(* IEC 61131-3 sources: daoli-st-library/DL_Algo (part 19) *)

(* ---- FB_DL_Q15BiquadFilter.st ---- *)
(*
  FB_DL_Q15BiquadFilter —— Q15 定点二阶 IIR 滤波：系数定点化、中间累加防溢出、移位饱和输出
  分类：DL_Algo | 复杂度：3 | 轮次：R86
  开源溯源：道莅原创（clean-room 自研，纯 IEC 61131-3 通用算法），无外部代码引用
  许可证：MIT

  职责：以直接 II 型转置（DF2T）结构实现二阶 IIR：y[n] = b0*x[n] + z1[n-1]；
        z1[n] = b1*x[n] - a1*y[n] + z2[n-1]；z2[n] = b2*x[n] - a2*y[n]。
        全部乘加在 DINT 内完成（Q15 × Q15 得 Q30），统一做「四舍五入右移 15 位 + Q15 饱和」，不调用任何外部库件。
  输入契约：arrCoef[0..4] = b0 / b1 / b2 / a1 / a2，均为 Q15 系数（±1.0 对应 ±32767）；
            iIn 为 Q15 输入；xReset 上升至真清历史；xEnable = FALSE 时清历史并输出 0。
  输出契约：iOut 为 Q15 输出；xOverflow 表示本拍发生了乘法累加或输出的饱和（信息级，可每拍重算）。
  边界：① 无除法、无开方，除零风险为零；② 所有移位用「乘 32768 / 除 32768」表达，避免方言 SHL/SHR 语义差异；
        ③ 定点饱和阈值 Q15_MAX / Q15_MIN 用 VAR CONSTANT 钉死；④ 零全局耦合、零物理地址、零库件依赖（R16）。
*)

FUNCTION_BLOCK FB_DL_Q15BiquadFilter
VAR_INPUT
    xEnable  : BOOL := TRUE;                              // 使能，FALSE 时清历史并输出零 [—] / Enable, false clears history
    xReset   : BOOL := FALSE;                             // 复位，真时清历史（单拍即可，无需沿） [—] / Reset, clears the history
    iIn      : INT  := 0;                                 // Q15 定点输入 [Q15] / The Q15 fixed point input
    arrCoef  : ARRAY[0..4] OF INT;                        // Q15 系数 b0/b1/b2/a1/a2 [Q15] / The Q15 coefficients
END_VAR
VAR_OUTPUT
    iOut      : INT;                                      // Q15 定点输出 [Q15] / The Q15 fixed point output
    xOverflow : BOOL;                                     // 本拍发生饱和（信息级） [—] / A saturation occurred this scan
END_VAR
VAR
    arrHist   : ARRAY[0..3] OF INT;                       // 历史：0=z1 1=z2 2=上拍输入 3=上拍输出 [Q15] / History slots
    diProd1   : DINT;                                     // 第一乘积项（Q30） [Q30] / The first product term
    diProd2   : DINT;                                     // 第二乘积项（Q30） [Q30] / The second product term
    diAcc     : DINT;                                     // 累加器（Q30） [Q30] / The Q30 accumulator
    diSh      : DINT;                                     // 四舍五入右移后的 Q15 暂存 [Q15] / The rounded Q15 stage
    diSum     : DINT;                                     // Q15 域饱和加法暂存 [Q15] / The Q15 domain saturating sum
    iNewZ1    : INT;                                      // 新的 z1 状态 [Q15] / The new z1 state
    iNewZ2    : INT;                                      // 新的 z2 状态 [Q15] / The new z2 state
    iSat      : INT;                                      // 饱和后的输出暂存 [Q15] / The saturated output stage
END_VAR
VAR CONSTANT
    Q15_MAX   : DINT := 32767;                            // Q15 上界 [-] / The Q15 upper bound
    Q15_MIN   : DINT := -32768;                           // Q15 下界 [-] / The Q15 lower bound
    DL_BQ_RND : DINT := 16384;                            // 右移 15 位的四舍五入偏置（2^14） [-] / The rounding bias
    DL_BQ_SC  : DINT := 32768;                            // Q15 定标因子（2^15） [-] / The Q15 scaling factor
    DL_BQ_Z   : DINT := 0;                                // 整型零常量 [Q15] / The integer zero constant
    DL_BQ_I0  : INT := 0;                                 // 整型零常量（INT 域） [Q15] / The integer zero constant in INT domain
    DL_BQ_I1  : INT := 1;                                 // 整型一常量（下标） [下标] / The integer one constant
    DL_BQ_I2  : INT := 2;                                 // 整型二常量（下标） [下标] / The integer two constant
    DL_BQ_I3  : INT := 3;                                 // 整型三常量（下标） [下标] / The integer three constant
    DL_BQ_I4  : INT := 4;                                 // 整型四常量（下标） [下标] / The integer four constant
END_VAR

// 段 1｜出口预置（本拍饱和标志每拍重算，属信息级）
xOverflow := FALSE;                                       // 饱和标志预置假 / preset the saturation flag false
iOut := DL_BQ_I0;                                         // 输出预置零 [Q15] / preset the output zero

// 段 2｜复位 / 失能闸：清全部历史并输出零（唯一复位路径）
IF xReset OR NOT xEnable THEN                             // 复位或失能 / reset asserted or disabled
    arrHist[DL_BQ_I0] := DL_BQ_I0;                        // z1 清零 [Q15] / clear z1
    arrHist[DL_BQ_I1] := DL_BQ_I0;                        // z2 清零 [Q15] / clear z2
    arrHist[DL_BQ_I2] := DL_BQ_I0;                        // 上拍输入清零 [Q15] / clear the previous input
    arrHist[DL_BQ_I3] := DL_BQ_I0;                        // 上拍输出清零 [Q15] / clear the previous output
    iOut := DL_BQ_I0;                                     // 输出零 [Q15] / output zero
    xOverflow := FALSE;                                   // 清饱和标志 [—] / clear the saturation flag
ELSE
    // 段 3｜y[n] = b0*x[n] + z1[n-1]（两项之和界内可证：|b0*x| <= 1.073e9，|z1*2^15| <= 1.073e9）
    diProd1 := INT_TO_DINT(arrCoef[DL_BQ_I0]) * INT_TO_DINT(iIn);          // b0*x [Q30] / b0 times x
    diProd2 := INT_TO_DINT(arrHist[DL_BQ_I0]) * DL_BQ_SC;                  // z1 左移 15 位 [Q30] / z1 scaled to Q30
    diAcc := diProd1 + diProd2;                                            // 两项求和 [Q30] / sum the two terms
    IF diAcc >= DL_BQ_Z THEN                                               // 非负做加偏置舍入 / non negative rounding
        diSh := (diAcc + DL_BQ_RND) / DL_BQ_SC;                            // 四舍五入右移 15 位 [Q15] / rounded shift right
    ELSE
        diSh := (diAcc - DL_BQ_RND) / DL_BQ_SC;                            // 负值做减偏置舍入 [Q15] / rounded shift right
    END_IF
    IF diSh > Q15_MAX THEN                                                 // 输出上越界 / the output exceeds the upper bound
        iSat := DINT_TO_INT(Q15_MAX);                                      // 饱和到 Q15_MAX [Q15] / saturate high
        xOverflow := TRUE;                                                 // 置饱和标志 [—] / raise the saturation flag
    ELSIF diSh < Q15_MIN THEN                                              // 输出下越界 / the output exceeds the lower bound
        iSat := DINT_TO_INT(Q15_MIN);                                      // 饱和到 Q15_MIN [Q15] / saturate low
        xOverflow := TRUE;                                                 // 置饱和标志 [—] / raise the saturation flag
    ELSE
        iSat := DINT_TO_INT(diSh);                                         // 界内直接转换 [Q15] / in range conversion
    END_IF
    iOut := iSat;                                                          // 本拍输出 [Q15] / the output of this scan

    // 段 4｜z1[n] = b1*x[n] - a1*y[n] + z2[n-1]（先算 Q30 两项差，再移位，再在 Q15 域饱和加 z2）
    diProd1 := INT_TO_DINT(arrCoef[DL_BQ_I1]) * INT_TO_DINT(iIn);          // b1*x [Q30] / b1 times x
    diProd2 := INT_TO_DINT(arrCoef[DL_BQ_I3]) * INT_TO_DINT(iSat);         // a1*y [Q30] / a1 times y
    diAcc := diProd1 - diProd2;                                            // 两项差（界内 |差| <= 2.147e9 可证） [Q30]
    IF diAcc >= DL_BQ_Z THEN                                               // 非负做加偏置舍入 / non negative rounding
        diSh := (diAcc + DL_BQ_RND) / DL_BQ_SC;                            // 四舍五入右移 15 位 [Q15] / rounded shift right
    ELSE
        diSh := (diAcc - DL_BQ_RND) / DL_BQ_SC;                            // 负值做减偏置舍入 [Q15] / rounded shift right
    END_IF
    diSum := diSh + INT_TO_DINT(arrHist[DL_BQ_I1]);                        // 加上 z2（|和| <= 98304 界内） [Q15] / add z2
    IF diSum > Q15_MAX THEN                                                // z1 上越界 / z1 exceeds the upper bound
        iNewZ1 := DINT_TO_INT(Q15_MAX);                                    // 饱和到 Q15_MAX [Q15] / saturate high
        xOverflow := TRUE;                                                 // 置饱和标志 [—] / raise the saturation flag
    ELSIF diSum < Q15_MIN THEN                                             // z1 下越界 / z1 exceeds the lower bound
        iNewZ1 := DINT_TO_INT(Q15_MIN);                                    // 饱和到 Q15_MIN [Q15] / saturate low
        xOverflow := TRUE;                                                 // 置饱和标志 [—] / raise the saturation flag
    ELSE
        iNewZ1 := DINT_TO_INT(diSum);                                      // 界内直接转换 [Q15] / in range conversion
    END_IF

    // 段 5｜z2[n] = b2*x[n] - a2*y[n]（同段 4 的判溢出 + 舍入 + 饱和口径）
    diProd1 := INT_TO_DINT(arrCoef[DL_BQ_I2]) * INT_TO_DINT(iIn);          // b2*x [Q30] / b2 times x
    diProd2 := INT_TO_DINT(arrCoef[DL_BQ_I4]) * INT_TO_DINT(iSat);         // a2*y [Q30] / a2 times y
    diAcc := diProd1 - diProd2;                                            // 两项差 [Q30] / the difference of the two terms
    IF diAcc >= DL_BQ_Z THEN                                               // 非负做加偏置舍入 / non negative rounding
        diSh := (diAcc + DL_BQ_RND) / DL_BQ_SC;                            // 四舍五入右移 15 位 [Q15] / rounded shift right
    ELSE
        diSh := (diAcc - DL_BQ_RND) / DL_BQ_SC;                            // 负值做减偏置舍入 [Q15] / rounded shift right
    END_IF
    IF diSh > Q15_MAX THEN                                                 // z2 上越界 / z2 exceeds the upper bound
        iNewZ2 := DINT_TO_INT(Q15_MAX);                                    // 饱和到 Q15_MAX [Q15] / saturate high
        xOverflow := TRUE;                                                 // 置饱和标志 [—] / raise the saturation flag
    ELSIF diSh < Q15_MIN THEN                                              // z2 下越界 / z2 exceeds the lower bound
        iNewZ2 := DINT_TO_INT(Q15_MIN);                                    // 饱和到 Q15_MIN [Q15] / saturate low
        xOverflow := TRUE;                                                 // 置饱和标志 [—] / raise the saturation flag
    ELSE
        iNewZ2 := DINT_TO_INT(diSh);                                       // 界内直接转换 [Q15] / in range conversion
    END_IF

    // 段 6｜状态统一提交（两段式：先算新值后写回，避免同拍读写串扰）
    arrHist[DL_BQ_I2] := iIn;                                             // 记录上拍输入 [Q15] / record the previous input
    arrHist[DL_BQ_I3] := iSat;                                            // 记录上拍输出 [Q15] / record the previous output
    arrHist[DL_BQ_I0] := iNewZ1;                                          // 提交新的 z1 [Q15] / commit z1
    arrHist[DL_BQ_I1] := iNewZ2;                                          // 提交新的 z2 [Q15] / commit z2
END_IF
END_FUNCTION_BLOCK

(* ---- FB_DL_QuantizeFilter.st ---- *)
(*==============================================================================
 * 组件名称 (Component)  : FB_DL_QuantizeFilter
 * 所属子库 (Sublibrary) : DL_Algo
 * 当前版本 (Version)    : 1.0.0
 * 兼容性   (Platform)   : CODESYS 3.5+ / TwinCAT 3 / 汇川 InoProShop / 施耐德 Machine Expert
 *                         仅依赖 Standard.library（ROUND / ABS），零厂商私有库
 * 功能描述 (Function)   : **量化取整 + 回差防抖**（有状态件）。
 *                         第一步量化：fQ := ROUND(fIn / fStep) × fStep（就近取整到步距倍数）；
 *                         第二步回差：仅当 |fQ - fOut| > fHyst 时才把 fOut 更新为 fQ，
 *                         否则保持。两步合起来解决「量化值在相邻两档之间反复跳」的现场顽症
 *                         （典型：0.5 单位步距的设定值显示与控制字抖动）。
 *                         与无状态取整 FC（FC_DL_QuantizeStep）的差别：那件每拍直接输出
 *                         量化值、无记忆；本件带上一档记忆与回差，切换次数显著下降。
 * 接口     (Interface)  : 输入 bEnable 使能、bReset 复位到当前量化值、fIn 采样输入 [EU]、
 *                         fStep 量化步距（必须 > 0） [EU]、fHyst 切换回差（>= 0） [EU]；
 *                         输出 fOut 量化并防抖后的输出 [EU]、fQuantized 原始量化值（诊断） [EU]、
 *                         bUpdated 本拍是否切换档位、bValid 输出有效、bError、uErrorId。
 * 边界     (Boundary)   : ① 属主边界：只做步距量化与回差防抖，不做死区保持（另件）、不做限速（另件）。
 *                         ② **除零防护（R4 硬要求）**：fStep 参与除法 fIn / fStep，
 *                         必须先判 fStep > 0，否则故障级 16#0009_0003，输出冻结。
 *                         fStep = 0 不允许「静默当直通」，否则调用方看不出配置错误。
 *                         ③ fHyst < 0 → 故障级 16#0009_0003（负回差等于放大抖动）。
 *                         ④ 非有限防御：fIn / fStep / fHyst 三个浮点入参逐一枚举。
 *                         ⑤ 取整一律用 ROUND（禁止 TRUNC(x)+1 这类手工进位）。
 *                         ⑥ 恢复路径：bEnable=FALSE 或 bReset=TRUE 解除故障态。
 *                         ⑦ 零全局耦合（无 GVL / VAR_EXTERNAL / 物理地址）。
 * 分工声明 (Scope)      : 与无状态 `FC_DL_QuantizeStep` 分工：单拍取整归那件、
 *                         带记忆的回差防抖归本件；与 `FB_DL_DeadbandFilter` 分工：
 *                         连续量死区归那件、离散档位回差归本件。
 * 来源标签 (Source Tag) : 原创实现（无外部代码引入）
 * 码表     (Codes)      : 16#0009_0000 无故障 / 16#0009_0002 入参非有限（故障级）/
 *                         16#0009_0003 步距或回差非法（故障级）/ 16#0009_0005 非法状态（故障级）。
 * 红线自检 (Redline)    : R1 ✓ 零 GVL/VAR_EXTERNAL ｜ R2 ✓ 零 %I/%Q/%M ｜ R3 ✓ 纯 IEC 61131-3
 *                         R4 ✓ 步距前置判零（除零防护）+ 三浮点入参非有限判 + ROUND 取整 ｜ R5 ✓ 声明逐行同行双语注释
 *                         R6 ✓ 四态 ENUM + CASE + ELSE 兜底 ｜ R7 N/A（无 TON / 边沿实例）
 * 修订历史 (Revision)   : 2026-11-23  v1.0.0  R77 首版（批次 B3 · 序号 15）
 * 验收向量 (Acceptance) : ① fStep=0.5, fHyst=0.2, fIn=1.24 → fQ=ROUND(2.48)×0.5=2×0.5=1.0，
 *                         |1.0 - fOut(初 0)|=1.0 > 0.2 → fOut=1.0, bUpdated=TRUE；
 *                         ② 随后 fIn=1.26 → fQ=ROUND(2.52)×0.5=3×0.5=1.5，|1.5-1.0|=0.5 > 0.2 → fOut=1.5；
 *                         ③ 随后 fIn=1.30 → fQ=1.5，|1.5-1.5|=0 <= 0.2 → fOut 保持 1.5, bUpdated=FALSE；
 *                         ④ fStep=0.0 → uErrorId=16#0009_0003，bError=TRUE（不静默直通）；
 *                         ⑤ fHyst=-0.1 → uErrorId=16#0009_0003，bError=TRUE。
 *==============================================================================*)

(*-----------------------------------------------------------------------------
 * 枚举: E_DL_QuantState（量化防抖状态机，归属 DL_Algo，与本件同文件，全库唯一属主）
 *----------------------------------------------------------------------------*)
TYPE E_DL_QuantState :
(
    eInit  := 0,    // 首扫 / 复位后：输出直取当前量化值 / First scan or after reset: output equals quantized value
    eRun   := 10,   // 运行态：量化 + 回差判定 / Running: quantize plus hysteresis decision
    eHold  := 20,   // 保持态：未使能，输出冻结 / Hold: disabled, output frozen
    eFault := 99    // 故障态：输出冻结，等待 bEnable 跌落或 bReset / Fault: frozen until cleared
);
END_TYPE

FUNCTION_BLOCK FB_DL_QuantizeFilter
VAR_INPUT
    bEnable : BOOL := FALSE;   // 使能，FALSE 冻结输出 / Enable, FALSE freezes output
    bReset  : BOOL := FALSE;   // 复位到当前量化值（单拍有效） / Reset to current quantized value, single scan
    fIn     : LREAL := 0.0;    // 采样输入 [EU] / Sampling input [EU]
    fStep   : LREAL := 1.0;    // 量化步距，必须 > 0 [EU] / Quantisation step, must be positive [EU]
    fHyst   : LREAL := 0.0;    // 切换回差，必须 >= 0 [EU] / Switching hysteresis, must be non-negative [EU]
END_VAR
VAR_OUTPUT
    fOut       : LREAL;   // 量化并防抖后的输出 [EU] / Quantised and debounced output [EU]
    fQuantized : LREAL;   // 原始量化值（诊断用） [EU] / Raw quantised value for diagnostics [EU]
    bUpdated   : BOOL;    // 本拍是否切换档位 [-] / Whether the output switched this scan
    bValid     : BOOL;    // 输出有效标志 [-] / Output valid flag
    bError     : BOOL;    // 故障标志，与 uErrorId 联动 [-] / Fault flag coupled with uErrorId
    uErrorId   : UDINT;   // 故障码，0 = 无故障 [-] / Error code, zero means healthy
END_VAR
VAR
    _bNonFin : BOOL;              // 入参非有限标志 [-] / Non-finite input flag
    _fRatio  : LREAL;             // 步距倍数（取整前） [-] / Step multiple before rounding
    eState   : E_DL_QuantState;   // 状态机当前状态 [-] / Current state
END_VAR
VAR CONSTANT
    DL_QTF_ZERO : LREAL := 0.0;   // 零基准（含非有限判零） [-] / Zero base including non-finite probe
END_VAR

(* —— 段 1：非有限防御（fIn / fStep / fHyst 三入参逐一枚举） —— *)
uErrorId := 16#0009_0000;                          // 预置无故障 / Preset healthy
_bNonFin := (fIn <> fIn) OR ((fIn - fIn) <> DL_QTF_ZERO);            // 输入非有限 / Input non-finite
_bNonFin := _bNonFin OR (fStep <> fStep) OR ((fStep - fStep) <> DL_QTF_ZERO);   // 步距非有限
_bNonFin := _bNonFin OR (fHyst <> fHyst) OR ((fHyst - fHyst) <> DL_QTF_ZERO);   // 回差非有限
IF _bNonFin THEN
    eState   := eFault;                            // 强制故障态 / Force fault state
    uErrorId := 16#0009_0002;                      // 故障级：入参非有限 / Fault: non-finite input
END_IF

(* —— 段 2：步距与回差域闸（步距必须严格正：它是除数；回差必须非负） —— *)
IF (fStep <= DL_QTF_ZERO) OR (fHyst < DL_QTF_ZERO) THEN
    eState   := eFault;                            // 参数非法进故障态 / Illegal parameter goes to fault
    uErrorId := 16#0009_0003;                      // 故障级：步距或回差非法 / Fault: illegal step or hysteresis
    fQuantized := DL_QTF_ZERO;                     // 诊断量回 0 / Diagnostic value zeroed
END_IF

(* —— 段 3：复位请求 → 回首扫 —— *)
IF bReset THEN
    eState := eInit;
END_IF

(* —— 段 4：状态派生 —— *)
IF NOT bEnable THEN
    eState := eHold;                               // 未使能：冻结 / Disabled: freeze
ELSIF eState = eFault THEN
    eState := eFault;                              // 故障态保持 / Fault holds
ELSIF eState = eInit THEN
    eState := eInit;                               // 首扫保持一拍 / Init holds one scan
ELSE
    eState := eRun;
END_IF

(* —— 段 5：主状态机（CASE 覆盖 + ELSE 兜底） —— *)
CASE eState OF

    eInit:
        _fRatio     := fIn / fStep;                // 步距倍数（fStep 已在段 2 判正） / Step multiple, step proven positive
        fQuantized  := ROUND(_fRatio) * fStep;     // 就近量化（禁止 TRUNC+1 手工进位） / Nearest quantisation
        fOut        := fQuantized;                 // 首拍直取量化值 / First scan adopts quantised value
        bUpdated    := TRUE;
        bValid      := TRUE;
        eState      := eRun;

    eRun:
        _fRatio    := fIn / fStep;                 // 步距倍数 / Step multiple
        fQuantized := ROUND(_fRatio) * fStep;      // 就近量化 / Nearest quantisation
        IF ABS(fQuantized - fOut) > fHyst THEN
            fOut     := fQuantized;                // 超出回差：切换档位 / Beyond hysteresis: switch
            bUpdated := TRUE;
        ELSE
            (* 回差内：保持原档位，避免相邻档反复跳变 / Inside hysteresis: hold current step *)
            bUpdated := FALSE;
        END_IF
        bValid := TRUE;

    eHold:
        (* 未使能：输出、量化诊断值、切换标志全部冻结 / Disabled: output, diagnostic and flag frozen *)
        bUpdated := FALSE;
        bValid   := FALSE;

    eFault:
        (* 故障态：输出冻结保持上拍值（不推 0，避免下游误判） / Fault: output frozen *)
        bUpdated := FALSE;
        bValid   := FALSE;

    ELSE
        eState     := eFault;
        bUpdated   := FALSE;
        bValid     := FALSE;
        fQuantized := DL_QTF_ZERO;
        uErrorId   := 16#0009_0005;                // 故障级：非法状态 / Fault: illegal state

END_CASE;

(* —— 段 6：出口映射（bError 与 uErrorId 同源；本件无信息级码） —— *)
bError := (uErrorId <> 16#0009_0000);

END_FUNCTION_BLOCK

(* ---- FB_DL_RampGenerator.st ---- *)
(*==============================================================================
 * 组件名称 (Component)  : FB_DL_RampGenerator
 * 所属子库 (Sublibrary) : DL_Algo
 * 当前版本 (Version)    : 1.0.1
 * 兼容性   (Platform)   : CODESYS 3.5 / TwinCAT 3 / 汇川 InoProShop / Machine Expert
 *                         仅依赖 Standard.library（LIMIT / MIN / ABS / SIGN），零厂商方言
 * 功能描述 (Function)   : 线性设定值斜坡发生器。把阶跃目标值变为按独立上升/下降
 *                         速率（EU/s）平滑逼近的斜坡输出，防止操作员大阶跃直接
 *                         冲击执行器。支持暂停保持（bHold 冻结当前值）与跟踪回投
 *                         （bTrack + fTrackValue 投切无扰动）。
 *                         斜率为 0 表示该方向冻结（保持输出，绝不直通，防误操作）。
 *                         到达判定以限幅后的实际输出为准，防止目标超量程时死等。
 * 开源溯源 (Origin)     : 原创实现。算法思想源自 IEC 61131-3 标准函数语义与
 *                         PLCopen Coding Guidelines 的周期安全约定，
 *                         未复制任何厂商私有库源码。
 * 本文件内含       : TYPE  E_DL_RampState（配套枚举，归属 DL_Algo）
 *                    FB    FB_DL_RampGenerator
 * 依赖     (Depends)    : 无 DL_ 内部依赖；Standard.library: LIMIT / MIN / ABS / SIGN
 * 红线自检 (Redline)    : R1 ✓ 零全局变量表与外部变量引用 ｜ R2 ✓ 零物理 IO 地址直写
 *                         R3 ✓ 纯 IEC 61131-3 ｜ R4 ✓ 速率/量程钳位+非有限值拒绝
 *                         R5 ✓ 全变量中英双语同行注释 ｜ R6 ✓ 六态 ENUM+CASE+ELSE
 *                         R7 N/A（无定时器/边沿实例）
 * 【边界披露 / Boundary disclosure】
 *   B1 速率 <= 0 视为非法：置 16#0002_0601 且该方向步长为 0（冻结），绝不直通。
 *   B2 目标非有限值（NaN 或幅值超 1.0E30）：本拍拒绝更新，保持上一拍输出。
 *   B3 rOutMin > rOutMax：自动对调并置 16#0002_0001，不中断扫描。
 *   B4 目标超量程不截断目标，仅限幅输出；到达判定用限幅后实际值，防死等。
 * 【验收向量 / Acceptance vectors】
 *   V1  fTarget 0→100，fRateUp=10 EU/s，tSampleTime=T#100MS → 每拍 +1.0 EU，
 *       10 s 后 fOut≈100、bDone=TRUE
 *   V2  fTarget 100→30，fRateDown=10 EU/s → 每拍 -1.0 EU、bMoving=TRUE
 *   V3  bHold=TRUE → fOut 冻结、状态 eHold；释放后继续逼近目标
 *   V4  fRateUp=0 → 16#0002_0601，向上移动冻结、fOut 保持
 *   V5  bTrack 一拍（fTrackValue=50）→ fOut=50，下一拍从 50 继续斜坡（无扰动）
 *   V6  rOutMin=100 > rOutMax=0 → 自动对调、16#0002_0001
 *   V7  fTarget=NaN → 16#0002_0004，fOut 保持上一拍值
 * 修订历史 (Revision)   :
 *   2026-11-15  v1.0.0  首版入库（Round 04 · Phase 3 · DL_Algo 批次）
 *   2026-11-15  v1.0.1  阶段五终审精修：首扫自动跟踪判据修复（bInit 判据
 *                       反向导致首扫不跟踪），对齐通用约定 0-6
 *============================================================================*)

(*-----------------------------------------------------------------------------
 * 枚举: E_DL_RampState（归属 DL_Algo，与 FB_DL_RampGenerator 同文件）
 * 含义: 斜坡状态机离散状态。数值步长留空位便于后续插态而不破坏已有工程。
 *----------------------------------------------------------------------------*)
TYPE E_DL_RampState :
(
    eIdle    := 0,    // 空闲态：未使能或等待评估，输出保持 / Idle state, output frozen
    eHold    := 10,   // 暂停保持态：操作员请求冻结当前输出 / Hold state, output frozen on operator request
    eRampUp  := 20,   // 上升斜坡态：按 fRateUpEff 步进逼近目标 / Ramping up with effective up rate
    eRampDown:= 30,   // 下降斜坡态：按 fRateDownEff 步进逼近目标 / Ramping down with effective down rate
    eDone    := 40,   // 到达态：输出与目标偏差在容差内 / Done state, deviation within tolerance
    eFault   := 99    // 故障兜底态：非法状态拦截，自动回空闲 / Fault fallback, auto recover to idle
);
END_TYPE

(*==============================================================================
 * 功能块: FB_DL_RampGenerator
 * 调用约定: 每个扫描周期无条件调用一次；bTrack 使能时输出立即跟随 fTrackValue。
 * 无状态泄漏: 全部状态驻留于实例私有 VAR，可多实例并行互不影响。
 * 速率披露: 输出相对目标的延迟 = 偏差量 / 对应方向速率（线性，非固定时间）。
 *============================================================================*)
FUNCTION_BLOCK FB_DL_RampGenerator
VAR_INPUT
    bEnable     : BOOL := FALSE;        // 使能标志，FALSE 时斜坡停止并保持输出 / Enable flag, FALSE stops ramp and holds output
    fTarget     : REAL := 0.0;          // 目标值 [EU]，可为任意有限值 / Target value [EU], any finite value
    fRateUp     : REAL := 10.0;         // 上升速率 [EU/s]，<=0 视为非法冻结 / Up rate [EU/s], <=0 illegal and frozen
    fRateDown   : REAL := 10.0;         // 下降速率 [EU/s]，<=0 视为非法冻结 / Down rate [EU/s], <=0 illegal and frozen
    bHold       : BOOL := FALSE;        // 暂停保持请求，TRUE 冻结在当前值 / Hold request, TRUE freezes at current value
    bTrack      : BOOL := FALSE;        // 跟踪使能，TRUE 时输出立即跟随 fTrackValue / Track enable, output follows fTrackValue instantly
    fTrackValue : REAL := 0.0;          // 跟踪值 [EU]，投切无扰动基准 / Track value [EU], bumpless transfer reference
    rOutMin     : REAL := -1.0E10;      // 输出下限 [EU]，大于上限时自动对调 / Output lower limit [EU], swapped if greater
    rOutMax     : REAL := 1.0E10;       // 输出上限 [EU]，小于下限时自动对调 / Output upper limit [EU], swapped if smaller
    tSampleTime : TIME := T#100MS;      // 采样周期 [s]，小于 10ms 钳位为 10ms / Sample time [s], clamped to 10ms minimum
END_VAR
VAR_OUTPUT
    fOut        : REAL;                 // 斜坡输出 [EU] / Ramp output [EU]
    bDone       : BOOL;                 // 到达目标标志：偏差在容差内 / Done flag, deviation within tolerance
    bMoving     : BOOL;                 // 斜坡进行中标志 / Ramp in progress flag
    fRemain     : REAL;                 // 距目标剩余量 [EU] = fTarget - fOut / Remaining amount to target [EU]
    bError      : BOOL;                 // 故障标志（瞬时，逐拍重算） / Fault flag, transient, recomputed every scan
    uErrorId    : UDINT;                // 故障码，0 = 无故障 / Error code, 0 = no error
END_VAR
VAR
    fRateUpEff  : REAL;                 // 钳位后的有效上升速率 [EU/s] / Effective clamped up rate [EU/s]
    fRateDownEff: REAL;                 // 钳位后的有效下降速率 [EU/s] / Effective clamped down rate [EU/s]
    fDt         : REAL;                 // 折算后的采样周期 [s] / Converted sample period [s]
    fDelta      : REAL;                 // 本拍目标与输出的偏差 [EU] / Deviation between target and output [EU]
    fStep       : REAL;                 // 本拍允许的最大步长 [EU] / Max step allowed this scan [EU]
    bTgtValid   : BOOL;                 // 目标为有限值的合法性标志 / Target finite validity flag
    bInit       : BOOL;                 // 首扫标志：首扫自动跟踪 fTrackValue / First scan flag, auto track on first scan
    eState      : E_DL_RampState;       // 主状态机当前状态 / Current state of the main state machine
END_VAR
VAR CONSTANT
    DL_RAMP_EPS     : REAL := 1.0E-6;   // 到达判定容差 [EU]，浮点差值比较 / Arrival tolerance [EU], float diff compare
    DL_RAMP_RATE_MAX: REAL := 1.0E10;   // 速率上限钳位 [EU/s]，防溢出 / Rate upper clamp [EU/s], overflow guard
END_VAR

(*------------------------------------------------------------------------------
 * 段 1｜公共参数处理（通用约定 0-1/0-2/0-3）：周期钳位、量程对调、故障码瞬时清零
 *      Common parameter handling: sample time clamp, limit swap, transient code reset
 *-----------------------------------------------------------------------------*)
uErrorId := 16#0000_0000;               // 故障码逐拍重算（瞬时语义） / Error code recomputed every scan
bError   := FALSE;                      // 故障标志逐拍重算 / Fault flag recomputed every scan

IF tSampleTime < T#10MS THEN
    fDt      := TIME_TO_REAL(T#10MS) / 1000.0; // 非法周期钳位为 10ms / Illegal period clamped to 10ms
    uErrorId := 16#0002_0002;           // 采样周期非法已钳位 / Sample time illegal, clamped
ELSE
    fDt      := TIME_TO_REAL(tSampleTime) / 1000.0; // 周期换算为秒 [s] / Period converted to seconds [s]
END_IF

IF rOutMin > rOutMax THEN
    fOut := LIMIT(rOutMax, fOut, rOutMin); // 对调后按新序限幅输出 / Clamp output with swapped limits
    uErrorId := 16#0002_0001;           // 参数越界已对调 / Limits out of order, swapped
ELSE
    fOut := LIMIT(rOutMin, fOut, rOutMax); // 正常序限幅输出 / Clamp output with normal limits
END_IF

(*------------------------------------------------------------------------------
 * 段 2｜速率钳位：<=0 非法（冻结方向），超上限钳位（边界 B1）
 *      Rate clamping: <=0 illegal (freeze direction), over-limit clamped
 *-----------------------------------------------------------------------------*)
IF fRateUp <= 0.0 THEN
    fRateUpEff := 0.0;                  // 非法速率冻结为 0，步长为 0 / Illegal rate frozen to zero step
    uErrorId   := 16#0002_0601;         // 速率非法已钳位 / Rate illegal, clamped
ELSIF fRateUp > DL_RAMP_RATE_MAX THEN
    fRateUpEff := DL_RAMP_RATE_MAX;     // 超上限钳位防溢出 / Over-limit clamped for overflow guard
    uErrorId   := 16#0002_0601;         // 速率非法已钳位 / Rate illegal, clamped
ELSE
    fRateUpEff := fRateUp;              // 合法速率直通 / Valid rate passed through
END_IF

IF fRateDown <= 0.0 THEN
    fRateDownEff := 0.0;                // 非法速率冻结为 0，步长为 0 / Illegal rate frozen to zero step
    uErrorId     := 16#0002_0601;       // 速率非法已钳位 / Rate illegal, clamped
ELSIF fRateDown > DL_RAMP_RATE_MAX THEN
    fRateDownEff := DL_RAMP_RATE_MAX;   // 超上限钳位防溢出 / Over-limit clamped for overflow guard
    uErrorId     := 16#0002_0601;       // 速率非法已钳位 / Rate illegal, clamped
ELSE
    fRateDownEff := fRateDown;          // 合法速率直通 / Valid rate passed through
END_IF

(*------------------------------------------------------------------------------
 * 段 3｜目标合法性判定（边界 B2）：非有限值本拍拒绝，保持上一拍目标行为
 *      Target validity: non-finite value rejected this scan, previous behavior kept
 *-----------------------------------------------------------------------------*)
bTgtValid := NOT (fTarget <> fTarget) AND (ABS(fTarget) <= 1.0E30); // NaN 判别 + 幅值防御 / NaN check plus magnitude guard
IF NOT bTgtValid THEN
    uErrorId := 16#0002_0004;           // 输入非有限值已拒绝 / Non-finite input rejected
END_IF

(*------------------------------------------------------------------------------
 * 段 4｜跟踪与首扫（通用约定 0-6）：投切无扰动，首扫自动跟踪 fTrackValue
 *      Tracking and first scan: bumpless transfer, first scan auto track
 *-----------------------------------------------------------------------------*)
IF bTrack OR (NOT bInit) THEN
    fOut   := LIMIT(rOutMin, fTrackValue, rOutMax); // 输出立即跟随跟踪值 / Output follows track value instantly
    eState := eIdle;                    // 回空闲重新评估方向 / Back to idle for direction re-evaluation
    bInit  := TRUE;                     // 首扫标志置位 / First scan flag set
END_IF

(*------------------------------------------------------------------------------
 * 段 5｜主状态机（红线 R6）：ENUM + CASE + ELSE 兜底
 *      Main state machine: ENUM + CASE with mandatory ELSE fallback
 *-----------------------------------------------------------------------------*)
fDelta := fTarget - fOut;               // 本拍偏差 [EU] / Deviation this scan [EU]

IF NOT bEnable THEN
    eState := eIdle;                    // 未使能：强制空闲、输出保持 / Disabled: force idle, output held
ELSE
    CASE eState OF

        eIdle:  // 空闲态：使能后按偏差方向选择迁移 / Idle: pick transition by deviation direction
            IF bTgtValid AND ABS(fDelta) > DL_RAMP_EPS THEN
                IF bHold THEN
                    eState := eHold;    // 保持请求优先 / Hold request has priority
                ELSIF fDelta > 0.0 THEN
                    eState := eRampUp;  // 目标在上方，进入上升 / Target above, ramp up
                ELSE
                    eState := eRampDown; // 目标在下方，进入下降 / Target below, ramp down
                END_IF
            ELSIF bTgtValid THEN
                eState := eDone;        // 已在容差内，直接到达 / Already within tolerance, done
            END_IF

        eHold:  // 暂停保持态：冻结输出直到释放 / Hold: freeze output until released
            IF NOT bHold THEN
                IF ABS(fDelta) <= DL_RAMP_EPS THEN
                    eState := eDone;    // 保持期间目标已到达 / Target reached during hold
                ELSIF fDelta > 0.0 THEN
                    eState := eRampUp;  // 释放后继续上升 / Resume ramp up after release
                ELSE
                    eState := eRampDown; // 释放后继续下降 / Resume ramp down after release
                END_IF
            END_IF

        eRampUp:  // 上升斜坡态：步长 = MIN(偏差, 速率*周期) / Ramp up: step = MIN(deviation, rate*period)
            IF ABS(fDelta) <= DL_RAMP_EPS THEN
                eState := eDone;        // 到达目标 / Target reached
            ELSIF fDelta < 0.0 THEN
                eState := eRampDown;    // 目标反转为下方 / Target switched below
            ELSIF bHold THEN
                eState := eHold;        // 保持请求 / Hold request
            ELSE
                fStep := MIN(fDelta, fRateUpEff * fDt); // 本拍步长 [EU] / Step this scan [EU]
                fOut  := fOut + fStep;  // 逐步逼近目标 / Step toward target
            END_IF

        eRampDown:  // 下降斜坡态：对称逻辑 / Ramp down: symmetric logic
            IF ABS(fDelta) <= DL_RAMP_EPS THEN
                eState := eDone;        // 到达目标 / Target reached
            ELSIF fDelta > 0.0 THEN
                eState := eRampUp;      // 目标反转为上方 / Target switched above
            ELSIF bHold THEN
                eState := eHold;        // 保持请求 / Hold request
            ELSE
                fStep := MIN(-fDelta, fRateDownEff * fDt); // 本拍步长 [EU] / Step this scan [EU]
                fOut  := fOut - fStep;  // 逐步逼近目标 / Step toward target
            END_IF

        eDone:  // 到达态：监视新目标 / Done: watch for new target
            IF bTgtValid AND ABS(fDelta) > DL_RAMP_EPS THEN
                IF bHold THEN
                    eState := eHold;    // 保持请求 / Hold request
                ELSIF fDelta > 0.0 THEN
                    eState := eRampUp;  // 新目标在上方 / New target above
                ELSE
                    eState := eRampDown; // 新目标在下方 / New target below
                END_IF
            END_IF

        eFault:  // 故障兜底态：无复位引脚，当拍回空闲重评，避免永久锁死 / Fault fallback: no reset pin, recover to idle
            eState := eIdle;            // 自动恢复空闲 / Auto recover to idle

        ELSE  // 非法状态拦截：任何未定义状态一律进故障态并置码 / Illegal state interception
            eState   := eFault;         // 强制故障态 / Force fault state
            uErrorId := 16#0002_0005;   // 非法状态兜底 / Illegal state fallback
            bError   := TRUE;           // 故障标志置位 / Fault flag set

    END_CASE;
END_IF

(*------------------------------------------------------------------------------
 * 段 6｜输出整形与状态引脚：限幅后实际值判定到达（边界 B4 防死等）
 *      Output shaping and status pins: arrival judged on clamped actual output
 *-----------------------------------------------------------------------------*)
IF rOutMin > rOutMax THEN
    fOut := LIMIT(rOutMax, fOut, rOutMin); // 对调序限幅（与段 1 一致） / Clamp with swapped order
ELSE
    fOut := LIMIT(rOutMin, fOut, rOutMax); // 正常序限幅 / Clamp with normal order
END_IF

fDelta  := fTarget - fOut;              // 限幅后重算偏差 [EU] / Deviation recomputed after clamping
fRemain := fDelta;                      // 距目标余量 [EU] / Remaining to target [EU]

bDone   := bEnable AND bTgtValid AND (ABS(fDelta) <= DL_RAMP_EPS); // 到达标志 / Done flag
bMoving := bEnable AND bTgtValid AND (NOT bHold)
           AND (ABS(fDelta) > DL_RAMP_EPS)
           AND ((eState = eRampUp) OR (eState = eRampDown));        // 斜坡进行中 / Ramp in progress
END_FUNCTION_BLOCK

(* ---- FB_DL_RateLimiter.st ---- *)
(*==============================================================================
 * 组件名称 (Component)  : FB_DL_RateLimiter
 * 所属子库 (Sublibrary) : DL_Algo
 * 当前版本 (Version)    : 1.0.0
 * 兼容性   (Platform)   : CODESYS 3.5 / TwinCAT 3 / 汇川 InoProShop / Machine Expert
 *                         仅依赖纯 IEC 61131-3 数学运算，零库依赖，零厂商方言
 * 功能描述 (Function)   : 变化率限制器（对应变化率限制语义）。输入阶跃时输出
 *                         以最大速率跟随，保护加热元件 / 执行器免受给定值阶跃
 *                         冲击；上升与下降速率独立可调，速率为 0 表示该方向不
 *                         限速直通（沿测量库惯例），负值非法按 0 处理并置码；
 *                         支持跟踪回投与限速进行中标志。
 * 开源溯源 (Origin)     : 原创实现。功能分类与参数域参考测量函数库中变化率
 *                         限制单元的公开语义描述，未复制任何厂商源码，
 *                         clean-room 重写。
 * 本文件内含       : TYPE  E_DL_RateState（配套枚举，归属 DL_Algo）
 *                    FB    FB_DL_RateLimiter
 * 依赖     (Depends)    : 无 DL_ 内部依赖；Standard.library 无实例依赖
 * 红线自检 (Redline)    : R1 ✓ 零全局变量表与外部变量引用 ｜ R2 ✓ 零物理 IO 地址直写
 *                         R3 ✓ 纯 IEC 61131-3 ｜ R4 ✓ 防除零+钳位+非有限值防御
 *                         R5 ✓ 全变量中英双语同行注释 ｜ R6 ✓ 五态 ENUM+CASE+ELSE
 *                         R7 ✓ 本块无定时器 / 边沿实例（无可刷新项，天然合规）
 * 修订历史 (Revision)   :
 *   2026-11-15  v1.0.0  首版入库 · Round 04 · Level 1 DL_Algo
 * 验收向量 (Acceptance) :
 *   V1 上升限速：fRateUp=10 EU/s, 输入阶跃 +100 → 输出每拍 +1 EU（100 ms 周期）
 *   V2 下降限速：fRateDown=5 EU/s, 输入阶跃 -100 → 输出每拍 -0.5 EU
 *   V3 零速率直通：fRateUp=0 → 上升方向立即跟随输入
 *   V4 到达直通：输出追上输入后 bLimiting=FALSE 且输出等于输入
 *   V5 跟踪：bTrack 置位 → 输出立即等于 fTrackValue
 *   V6 非有限值：输入写非法浮点 → 输出保持上一拍且码 0002_0004
 *============================================================================*)

(*-----------------------------------------------------------------------------
 * 枚举: E_DL_RateState（归属 DL_Algo，与 FB_DL_RateLimiter 同文件）
 * 含义: 变化率限制离散状态。数值步长留空位便于后续插态而不破坏已有工程。
 *----------------------------------------------------------------------------*)
TYPE E_DL_RateState :
(
    eIdle      := 0,   // 使能关：输出直通输入 / Idle: enable off, output follows input
    eFollow    := 10,  // 不限速直通：两方向均无需限速 / Follow: no rate limit needed in either direction
    eLimitUp   := 20,  // 上升限速：输出按最大上升速率逼近 / Limit up: output approaches at max rise rate
    eLimitDown := 30,  // 下降限速：输出按最大下降速率逼近 / Limit down: output approaches at max fall rate
    eFault     := 99   // 故障兜底态：非法状态进入，输出保持 / Fault fallback: illegal state, output held
);
END_TYPE

(*==============================================================================
 * 功能块: FB_DL_RateLimiter
 * 调用约定: 每个扫描周期无条件调用一次；采样周期引脚按子库通用约定配置。
 * 无状态泄漏: 全部状态驻留于实例私有 VAR，零全局引用，可多实例并行。
 * 工程披露: 输出变量自身即斜坡历史状态，不另设历史缓冲；实际变化率按本拍
 *           输出增量除以采样周期计算，供 HMI 趋势与诊断。
 *============================================================================*)
FUNCTION_BLOCK FB_DL_RateLimiter
VAR_INPUT
    bEnable     : BOOL := FALSE;      // 总使能，FALSE 时输出直通输入 / Master enable, FALSE passes input through
    fIn         : REAL := 0.0;        // 输入信号 [EU] / Input signal in engineering units
    fRateUp     : REAL := 0.0;        // 最大上升速率 [EU/s]，0 = 不限 / Max rising rate, 0 = unlimited
    fRateDown   : REAL := 0.0;        // 最大下降速率 [EU/s]，0 = 不限 / Max falling rate, 0 = unlimited
    bTrack      : BOOL := FALSE;      // 跟踪使能，TRUE 时输出立即跟随跟踪值 / Track enable, output follows track value
    fTrackValue : REAL := 0.0;        // 跟踪值 [EU]，用于无扰投切 / Track value for bumpless transfer
    tSampleTime : TIME := T#100MS;    // 采样周期，按子库通用约定 / Sample period per sublibrary convention
END_VAR
VAR_OUTPUT
    fOut        : REAL;               // 限速后输出 [EU] / Rate-limited output in engineering units
    bLimiting   : BOOL;               // 限速进行中标志 / Rate limiting in progress flag
    fRateActual : REAL;               // 本拍实际变化率 [EU/s] / Actual rate of change this cycle
    bError      : BOOL;               // 故障标志 / Fault flag
    uErrorId    : UDINT;              // 故障码，0 = 无故障 / Error code, 0 = no error
END_VAR
VAR
    eState      : E_DL_RateState;     // 主状态机当前状态 / Current state of the state machine
    bInit       : BOOL := FALSE;      // 首扫初始化标志 / First-scan init flag
    fDt         : REAL;               // 生效采样周期 [s] / Effective sample period in seconds
    fRateUpEff  : REAL;               // 钳位后的有效上升速率 [EU/s] / Clamped effective rise rate
    fRateDownEff: REAL;               // 钳位后的有效下降速率 [EU/s] / Clamped effective fall rate
    fDelta      : REAL;               // 输入与输出的差值 [EU] / Difference between input and output
    fStepMax    : REAL;               // 本拍允许的最大步进 [EU] / Maximum allowed step this cycle
    fStepApply  : REAL;               // 本拍实际施加步进 [EU] / Actually applied step this cycle
    fOutBefore  : REAL;               // 本拍更新前的输出 [EU] / Output before this cycle update
    bNonFinite  : BOOL;               // 本拍输入非有限值标志 / Non-finite input flag of this cycle
END_VAR

(*------------------------------------------------------------------------------
 * 段 1｜参数钳位与公共防御（不中断扫描）
 *      Parameter clamping and common defenses, never stops the scan
 *-----------------------------------------------------------------------------*)
bError   := FALSE;                    // 每拍重算故障标志 / Recompute fault flag every cycle
uErrorId := 16#0002_0000;             // 每拍重算故障码 / Recompute error code every cycle
bLimiting := FALSE;                   // 限速标志每拍重算 / Limiting flag recomputed every cycle
bNonFinite := FALSE;                  // 非有限值标志每拍重算 / Non-finite flag recomputed every cycle

IF tSampleTime < T#10MS THEN
    fDt := 0.01;                      // 采样周期非法钳位为 0.01 s / Illegal sample period clamped to 0.01 s
    uErrorId := 16#0002_0002;         // 公共码：采样周期已钳位 / Common code: sample period clamped
ELSE
    fDt := TIME_TO_REAL(tSampleTime) / 1000.0;  // 采样周期换算为秒 [s] / Sample period in seconds
END_IF

(* 速率防御：负值非法按 0（不限速）处理并置码，正值直通 *)
(* Rate defense: negative treated as 0 (unlimited) with code, positive passed *)
IF fRateUp < 0.0 THEN
    fRateUpEff := 0.0;                // 负上升速率按 0 处理 / Negative rise rate treated as zero
    uErrorId := 16#0002_0001;         // 公共码：参数越界已钳位 / Common code: parameter clamped
ELSE
    fRateUpEff := fRateUp;            // 合法上升速率直通 / Valid rise rate passed
END_IF
IF fRateDown < 0.0 THEN
    fRateDownEff := 0.0;              // 负下降速率按 0 处理 / Negative fall rate treated as zero
    uErrorId := 16#0002_0001;         // 公共码：参数越界已钳位 / Common code: parameter clamped
ELSE
    fRateDownEff := fRateDown;        // 合法下降速率直通 / Valid fall rate passed
END_IF

(* 输入非有限值防御：非法浮点拒绝本拍更新，保持上一拍输出 *)
(* Non-finite defense: reject this cycle, hold previous output *)
IF (fIn <> fIn) OR (ABS(fIn) > 1.0E30)
   OR (fTrackValue <> fTrackValue) OR (ABS(fTrackValue) > 1.0E30) THEN
    bNonFinite := TRUE;               // 置非有限值标志 / Set non-finite flag
    bError   := TRUE;                 // 置故障标志 / Set fault flag
    uErrorId := 16#0002_0004;         // 公共码：输入非有限值已拒绝 / Common code: non-finite rejected
END_IF

(*------------------------------------------------------------------------------
 * 段 2｜早退：使能关 / 非有限值 / 跟踪，输出直通或保持，状态机旁路
 *      Early exits: disable, non-finite, track; output passes or holds
 *-----------------------------------------------------------------------------*)
IF bNonFinite THEN
    RETURN;                           // 保持上一拍输出与状态 / Hold previous output and state
END_IF

IF NOT bEnable THEN
    eState := eIdle;                  // 强制回空闲态 / Force idle state
    fOut   := fIn;                    // 输出直通输入 / Output passes input through
    fRateActual := 0.0;               // 直通拍变化率为 0 / Zero rate on pass-through cycle
    bInit  := FALSE;                  // 复位首扫标志以便重使能时同步 / Reset init flag for resync
    RETURN;                           // 本拍结束 / End of this cycle
END_IF

IF bTrack OR (NOT bInit) THEN
    (* 跟踪回投 / 首扫初始化：输出立即同步，杜绝上电阶跃冲击 *)
    (* Track / first-scan init: output synchronized immediately, no power-up step *)
    IF bTrack THEN
        fOut := fTrackValue;          // 输出立即跟随跟踪值 / Output follows track value
    ELSE
        fOut := fIn;                  // 首扫输出直通输入 / First-scan output passes input
    END_IF
    eState := eFollow;                // 状态回直通态 / State back to follow
    fRateActual := 0.0;               // 同步拍变化率为 0 / Zero rate on sync cycle
    bInit  := TRUE;                   // 置首扫完成标志 / Set first-scan done flag
    RETURN;                           // 本拍结束 / End of this cycle
END_IF

(*------------------------------------------------------------------------------
 * 段 3｜限速需求判定：差值方向与有效速率共同决定本拍状态
 *      Limit demand: direction and effective rates decide this cycle state
 *-----------------------------------------------------------------------------*)
fDelta := fIn - fOut;                 // 输入与输出差值 [EU] / Input minus output difference
fOutBefore := fOut;                   // 记录更新前输出用于变化率计算 / Record output before update

IF fDelta > 0.0 THEN
    (* 上升需求：速率 0 直通，否则按最大上升步进逼近 *)
    (* Rise demand: zero rate passes through, else approach at max rise step *)
    IF fRateUpEff > 0.0 THEN
        eState := eLimitUp;           // 进上升限速态 / Enter rise-limit state
    ELSE
        eState := eFollow;            // 不限速直通 / Unlimited follow
    END_IF
ELSIF fDelta < 0.0 THEN
    (* 下降需求：速率 0 直通，否则按最大下降步进逼近 *)
    (* Fall demand: zero rate passes through, else approach at max fall step *)
    IF fRateDownEff > 0.0 THEN
        eState := eLimitDown;         // 进下降限速态 / Enter fall-limit state
    ELSE
        eState := eFollow;            // 不限速直通 / Unlimited follow
    END_IF
ELSE
    eState := eFollow;                // 已到达：直通 / Reached: follow
END_IF

(*------------------------------------------------------------------------------
 * 段 4｜主状态机（红线 R6）：ENUM + CASE + ELSE 兜底
 *      Main state machine: ENUM + CASE with mandatory ELSE fallback
 *-----------------------------------------------------------------------------*)
CASE eState OF

    eIdle:
        (* 空闲态已在早退段处理；本分支仅做迁移防御 *)
        (* Idle handled in early exit; this branch only guards transfers *)
        fOut := fIn;                  // 直通输出 / Pass-through output
        fRateActual := 0.0;           // 变化率为 0 / Zero rate

    eFollow:
        (* 不限速直通：输出立即等于输入 *)
        (* Unlimited follow: output equals input immediately *)
        fOut := fIn;                  // 直通输出 / Pass-through output
        fRateActual := fDelta / fDt;  // 本拍实际变化率 [EU/s] / Actual rate this cycle

    eLimitUp:
        (* 上升限速：步进 = MIN(|差值|, 速率*dt)，方向取差值符号 *)
        (* Rise limit: step = MIN(|delta|, rate*dt) in delta direction *)
        fStepMax   := fRateUpEff * fDt;                             // 最大步进 [EU] / Maximum step
        fStepApply := MIN(ABS(fDelta), fStepMax) * 1.0;             // 施加步进 [EU] / Applied step
        fOut       := fOutBefore + fStepApply;                      // 输出推进 / Output advanced
        bLimiting  := (ABS(fDelta) > fStepMax);                     // 限速进行中 / Limiting in progress
        fRateActual := fStepApply / fDt;                            // 本拍实际变化率 / Actual rate this cycle

    eLimitDown:
        (* 下降限速：步进取负方向 *)
        (* Fall limit: step taken in negative direction *)
        fStepMax   := fRateDownEff * fDt;                           // 最大步进 [EU] / Maximum step
        fStepApply := MIN(ABS(fDelta), fStepMax) * (-1.0);          // 施加步进 [EU] / Applied step
        fOut       := fOutBefore + fStepApply;                      // 输出推进 / Output advanced
        bLimiting  := (ABS(fDelta) > fStepMax);                     // 限速进行中 / Limiting in progress
        fRateActual := fStepApply / fDt;                            // 本拍实际变化率 / Actual rate this cycle

    eFault:
        (* 故障兜底态：输出保持上一拍值 *)
        (* Fault fallback: output holds previous value *)
        fOut := fOutBefore;           // 输出保持 / Output held
        fRateActual := 0.0;           // 变化率为 0 / Zero rate

    ELSE
        (* 非法状态拦截：任何未定义状态一律进故障兜底，不做隐式恢复 *)
        (* Illegal state interception: any undefined state goes to fault fallback *)
        eState   := eFault;           // 进故障态 / Enter fault state
        bError   := TRUE;             // 置故障标志 / Set fault flag
        uErrorId := 16#0002_0005;     // 非法状态兜底码 / Illegal state fallback code
        fOut     := fOutBefore;       // 输出保持 / Output held
        fRateActual := 0.0;           // 变化率为 0 / Zero rate
END_CASE;
END_FUNCTION_BLOCK

(* ---- FB_DL_RateOfChangeFilter.st ---- *)
(*==============================================================================
 * 组件名称 (Component)  : FB_DL_RateOfChangeFilter
 * 所属子库 (Sublibrary) : DL_Algo
 * 当前版本 (Version)    : 1.0.0
 * 兼容性   (Platform)   : CODESYS 3.5+ / TwinCAT 3 / 汇川 InoProShop / 施耐德 Machine Expert
 *                         仅依赖 Standard.library（ABS / MIN / MAX / TIME_TO_REAL），零厂商私有库
 * 功能描述 (Function)   : 变化率限幅滤波（斜坡限速）。每周期允许的最大增量
 *                         fMaxStep = fMaxRate × fDt（fDt 由 tSampleTime 显式给定），
 *                         输出增量被钳制在 ±fMaxStep 内：
 *                           fOut := fOut + LIMIT(fIn - fOut, -fMaxStep, +fMaxStep)
 *                         作用：抑制阶跃冲击（传感器跳变、通信坏包、量程切换瞬态），
 *                         保护下游执行机构与 PID 微分项，同时不引入一阶滞后（稳态无误差）。
 *                         与低通滤波的本质差别：本件**稳态增益恒为 1、无相位滞后**，
 *                         只在斜率上设限；阶跃会被摊成斜坡而非指数逼近。
 * 接口     (Interface)  : 输入 bEnable 使能、bReset 复位输出到当前输入、fIn 采样输入 [EU]、
 *                         fMaxRate 最大变化率 [EU/s]、tSampleTime 采样周期 [s]；
 *                         输出 fOut 限幅输出 [EU]、fMaxStep 本拍允许最大增量 [EU]、
 *                         bLimited 本拍是否发生限幅、bValid 输出有效、bError、uErrorId。
 * 边界     (Boundary)   : ① 属主边界：只做斜率限幅，不做低通 / 中值 / 死区（另件）。
 *                         ② 非有限防御覆盖 **fIn 与 fMaxRate 两个浮点入参**（漏一个即该判据静默失效）。
 *                         ③ 除零/非法参数防护：fMaxRate <= 0 → 故障级 16#0005_0003（不静默当 0 处理，
 *                         否则输出会被永久冻结而现场看不出原因）；tSampleTime < 10MS →
 *                         钳到 10MS 并置信息码 16#0005_0001。
 *                         ④ 复位语义：bReset=TRUE 当拍 fOut := fIn 且不计限幅，恢复无爬升。
 *                         ⑤ 零全局耦合（无 GVL / VAR_EXTERNAL / 物理地址）。
 * 分工声明 (Scope)      : 与 `FB_DL_LowPassFilter` 分工：一阶惯性与相位滞后归那件、
 *                         纯斜率限幅归本件；与 `FB_DL_GatedUpdateFilter` 分工：门控归那件。
 * 来源标签 (Source Tag) : 原创实现（无外部代码引入）
 * 码表     (Codes)      : 16#0005_0000 无故障 / 16#0005_0001 采样周期非法已钳位（信息级）/
 *                         16#0005_0002 输入非有限（故障级）/ 16#0005_0003 变化率非法（故障级）/
 *                         16#0005_0005 非法状态（故障级）。
 * 红线自检 (Redline)    : R1 ✓ 零 GVL/VAR_EXTERNAL ｜ R2 ✓ 零 %I/%Q/%M ｜ R3 ✓ 纯 IEC 61131-3
 *                         R4 ✓ 双浮点入参非有限判 + 变化率域闸 + 周期下限钳位 ｜ R5 ✓ 声明逐行同行双语注释
 *                         R6 ✓ 四态 ENUM + CASE + ELSE 兜底 ｜ R7 N/A（无 TON / 边沿实例）
 * 修订历史 (Revision)   : 2026-11-23  v1.0.0  R77 首版（批次 B3 · 序号 11）
 * 验收向量 (Acceptance) : ① fMaxRate=10, tSampleTime=T#100MS（fDt=0.1s）→ fMaxStep=1.0，
 *                         阶跃 0→100：第 1 拍 fOut=1.0、第 2 拍 fOut=2.0，bLimited=TRUE；
 *                         ② 稳态后 fIn 恒 100 → fOut 追到 100.0 时 bLimited=FALSE，无稳态误差；
 *                         ③ fMaxRate=0 → uErrorId=16#0005_0003，bError=TRUE，fOut 冻结；
 *                         ④ tSampleTime=T#1MS → 钳到 0.01s，uErrorId=16#0005_0001（不置 bError）；
 *                         ⑤ bReset=TRUE 一拍 → fOut 立即等于 fIn。
 *==============================================================================*)

(*-----------------------------------------------------------------------------
 * 枚举: E_DL_RocState（变化率限幅状态机，归属 DL_Algo，与本件同文件，全库唯一属主）
 *----------------------------------------------------------------------------*)
TYPE E_DL_RocState :
(
    eInit  := 0,    // 首扫 / 复位后：输出直取输入 / First scan or after reset: output follows input
    eRun   := 10,   // 运行态：按 fMaxStep 限幅 / Running: rate-limited stepping
    eHold  := 20,   // 保持态：未使能，输出冻结 / Hold: disabled, output frozen
    eFault := 99    // 故障态：输出冻结，等待 bEnable 跌落或 bReset / Fault: frozen until cleared
);
END_TYPE

FUNCTION_BLOCK FB_DL_RateOfChangeFilter
VAR_INPUT
    bEnable     : BOOL := FALSE;     // 使能，FALSE 冻结输出 / Enable, FALSE freezes output
    bReset      : BOOL := FALSE;     // 复位到当前输入（单拍有效） / Reset to current input, single scan
    fIn         : LREAL := 0.0;      // 采样输入 [EU] / Sampling input [EU]
    fMaxRate    : LREAL := 1.0;      // 最大变化率，必须 > 0 [EU/s] / Max rate of change, must be positive [EU/s]
    tSampleTime : TIME := T#100MS;   // 采样周期 [s]，小于 10ms 钳位 / Sampling period, clamped to 10ms
END_VAR
VAR_OUTPUT
    fOut     : LREAL;   // 限幅输出 [EU] / Rate-limited output [EU]
    fMaxStep : LREAL;   // 本拍允许最大增量 [EU] / Maximum allowed step this scan [EU]
    bLimited : BOOL;    // 本拍是否发生限幅 [-] / Whether limiting occurred this scan
    bValid   : BOOL;    // 输出有效标志 [-] / Output valid flag
    bError   : BOOL;    // 故障标志，与 uErrorId 联动 [-] / Fault flag coupled with uErrorId
    uErrorId : UDINT;   // 故障码，0 = 无故障 [-] / Error code, zero means healthy
END_VAR
VAR
    _fDt      : LREAL;         // 生效采样周期秒值 [s] / Effective sampling period in seconds
    _fDelta   : LREAL;         // 输入与输出的偏差 [EU] / Deviation between input and output
    _fStep    : LREAL;         // 本拍实际步进（已钳位） [EU] / Actual clamped step [EU]
    _bNonFin  : BOOL;          // 入参非有限标志 [-] / Non-finite input flag
    eState    : E_DL_RocState; // 状态机当前状态 [-] / Current state
END_VAR
VAR CONSTANT
    DL_ROC_DT_MIN  : LREAL := 0.01;     // 采样周期防御下限 [s] / Defensive sampling period floor [s]
    DL_ROC_ZERO    : LREAL := 0.0;      // 零基准（含非有限判零） [-] / Zero base including non-finite probe
    DL_ROC_MS      : LREAL := 1000.0;   // 毫秒转秒因子 [ms/s] / Milliseconds per second
END_VAR

(* —— 段 1：采样周期域闸（不中断扫描，只钳位并置信息码） —— *)
uErrorId := 16#0005_0000;                          // 预置无故障 / Preset healthy
IF tSampleTime < T#10MS THEN
    _fDt     := DL_ROC_DT_MIN;                     // 周期过小钳位 / Too small period clamped
    uErrorId := 16#0005_0001;                      // 信息级：采样周期已钳位 / Info: period clamped
ELSE
    _fDt := TIME_TO_REAL(tSampleTime) / DL_ROC_MS; // TIME 换算秒值 / Convert to seconds
END_IF

(* —— 段 2：非有限防御（fIn 与 fMaxRate 逐一枚举，禁止漏闸） —— *)
_bNonFin := (fIn <> fIn) OR ((fIn - fIn) <> DL_ROC_ZERO);            // 输入非有限 / Input non-finite
_bNonFin := _bNonFin OR (fMaxRate <> fMaxRate) OR ((fMaxRate - fMaxRate) <> DL_ROC_ZERO);  // 变化率非有限
IF _bNonFin THEN
    eState   := eFault;                            // 强制故障态 / Force fault state
    uErrorId := 16#0005_0002;                      // 故障级：入参非有限 / Fault: non-finite input
END_IF

(* —— 段 3：变化率域闸（必须严格为正，否则限幅无意义且输出会被永久冻结） —— *)
IF fMaxRate <= DL_ROC_ZERO THEN
    eState   := eFault;                            // 参数非法进故障态 / Illegal parameter goes to fault
    uErrorId := 16#0005_0003;                      // 故障级：变化率非法 / Fault: illegal rate
    fMaxStep := DL_ROC_ZERO;                       // 步长出口回 0（诊断量仍可读） / Step outlet zeroed
END_IF

(* —— 段 4：复位请求 → 回首扫 —— *)
IF bReset THEN
    eState := eInit;
END_IF

(* —— 段 5：状态派生 —— *)
IF NOT bEnable THEN
    eState := eHold;                               // 未使能：冻结 / Disabled: freeze
ELSIF eState = eFault THEN
    eState := eFault;                              // 故障态保持 / Fault holds
ELSIF eState = eInit THEN
    eState := eInit;                               // 首扫保持一拍 / Init holds one scan
ELSE
    eState := eRun;
END_IF

(* —— 段 6：主状态机（CASE 覆盖 + ELSE 兜底） —— *)
CASE eState OF

    eInit:
        fOut     := fIn;                           // 首拍直取输入，无历史瞬态 / First scan follows input
        fMaxStep := fMaxRate * _fDt;               // 步长按当前参数计算 / Step from current parameters
        bLimited := FALSE;
        bValid   := TRUE;
        eState   := eRun;

    eRun:
        fMaxStep := fMaxRate * _fDt;               // 本拍允许最大增量 [EU] / Maximum step this scan
        _fDelta  := fIn - fOut;                    // 偏差 / Deviation
        IF _fDelta > fMaxStep THEN
            _fStep   := fMaxStep;                  // 正向限幅 / Positive limiting
            bLimited := TRUE;
        ELSIF _fDelta < (DL_ROC_ZERO - fMaxStep) THEN
            _fStep   := DL_ROC_ZERO - fMaxStep;    // 负向限幅 / Negative limiting
            bLimited := TRUE;
        ELSE
            _fStep   := _fDelta;                   // 未超限：直接跟上（稳态无误差） / Within limit: track directly
            bLimited := FALSE;
        END_IF
        fOut   := fOut + _fStep;                   // 斜坡推进 / Ramp forward
        bValid := TRUE;

    eHold:
        (* 未使能：输出与步长诊断量保持上拍值 / Disabled: output and step diagnostics frozen *)
        bValid := FALSE;

    eFault:
        (* 故障态：输出冻结保持上拍值（不推 0，避免下游误判为真实零） / Fault: output frozen *)
        bValid := FALSE;

    ELSE
        eState   := eFault;
        bValid   := FALSE;
        fMaxStep := DL_ROC_ZERO;
        uErrorId := 16#0005_0005;                  // 故障级：非法状态 / Fault: illegal state

END_CASE;

(* —— 段 7：出口结果复检（非有限兜底，名实双出口） —— *)
IF (fOut <> fOut) OR ((fOut - fOut) <> DL_ROC_ZERO) THEN
    eState   := eFault;                            // 结果异常进故障态 / Abnormal result goes to fault
    bValid   := FALSE;
    uErrorId := 16#0005_0002;                      // 故障级码 / Fault-level code
END_IF
bError := (uErrorId <> 16#0005_0000) AND (uErrorId <> 16#0005_0001);   // 信息级不置 bError / Info level excluded

END_FUNCTION_BLOCK

(* ---- FB_DL_RatioController.st ---- *)
(*
    FB_DL_RatioController —— 比值控制站
    ------------------------------------------------------------------
    分类      : DL_Algo / ProcessControl
    前缀      : FB_DL_
    版本      : 1.0.0
    溯源      : 比值控制为公开过程控制通用结构（从动给定 = 主动流量 × 比率 + 偏置）；
                本件只借「参数域约束」的组织方式，低限切安全给定、迟滞式的状态迁移、
                斜率限制、兜底纪律与码位 100% 自有；clean-room 重写，未复制任何
                闭源厂商源码，参考实现仅限 MIT/Apache 许可
    平台      : 纯 IEC 61131-3，CODESYS V3.5+ / TwinCAT 3 / InoProShop 通用
    作者      : 道莅代码库 · PLC编程专家（R19）
    ------------------------------------------------------------------
    功能说明  : 从动流量给定 = 主动流量 × 比率 + 偏置。核心防御是「主动流量低限保护」：
                主动流量接近 0 时按比例算出的从动给定也趋 0，操作工看到「两个流量都归零」，
                真正的故障源（主动侧断料）被掩盖——本件在低限以下直接切到安全给定并置
                bMasterLow。其余防御：① 比率域与输出域自相矛盾即故障级 2811（区间不存在）；
                ② 比率越窗只钳位并置信息码（超窗是「待调整」而非故障）；
                ③ 斜率限制首拍 fStep = 0，绝不用 0 除；④ 输出双侧钳位（只做单侧是常见缺陷）；
                ⑤ 输入非有限时给定保持末次有效值——切 0 会直接停料；
                ⑥ 状态机 CASE 含 ELSE 兜底，非法状态回 eIdle 并保持末值。
                职责边界：本件不算 PID（环路闭合归 FB_DL_PidController），只出给定。
    错误码    : 16#0002_2801 比率被限幅 / 主动流量低于低限已切安全给定——信息级，正常防御
                16#0002_2802 预留禁用（信息级，不得挪用）
                16#0002_2810 输入非有限或斜率/采样参数非法——故障级，给定保持末次有效
                16#0002_2811 限值区间自相矛盾（比率域或输出域非法）——故障级，给定保持末次有效
                16#0002_2812 状态机落 ELSE 兜底（非法状态）——故障级，回 eIdle 并保持末值
    码位总账  : 16#0002_2801 用 / 16#0002_2802 预留 ｜ 16#0002_2810 用 / 16#0002_2811 用 / 16#0002_2812 用
    状态机    : E_DL_RatioState（eIdle / eRunning / eMasterLow / eFault）四态，CASE 含 ELSE 兜底，
                ELSE 分支回 eIdle 并置故障级 2812；失能无条件回 eIdle。
    采样约定  : fbTrigReset 在本体首部无条件刷新；斜率步长由 tSampleTime 引脚换算，
                首拍 fLastSp 未建立时 fStep 取 0（不做除零），故给定不会突变。
    修订记录  : 2026-11-16 v1.0.0 首次入库（R19）
*)

(*
    枚举 : E_DL_RatioState —— 比值站状态（本文件为全库唯一属主）
*)
TYPE E_DL_RatioState :
(
    eIdle      := 0,                          // 空闲：未使能，输出停在限幅下限 / idle, disabled, output parked at the lower bound
    eRunning   := 1,                          // 运行：按比率跟踪主动流量 / running, tracking the master flow by ratio
    eMasterLow := 2,                          // 主动低限：给定已切安全值 / master low, setpoint switched to the safe value
    eFault     := 3                           // 故障：给定保持末次有效值 / fault, setpoint holds the last valid value
);
END_TYPE

FUNCTION_BLOCK FB_DL_RatioController
VAR_INPUT
    bEnable         : BOOL;                   // 使能，FALSE 回 eIdle 并输出限幅下限 / enable, FALSE returns to eIdle and outputs the lower bound
    bReset          : BOOL;                   // 复位，上升沿清限幅锁存与斜率状态 / reset, rising edge clears the clamp latches and the ramp state
    fMasterFlow     : REAL := 0.0;            // 主动流量测量值 [m3/h]，范围 0.0~1.0E6 / measured master flow [m3/h], range 0.0~1.0E6
    fRatio          : REAL := 1.0;            // 比率 [无量纲]，范围 fRatioMin~fRatioMax / ratio [dimensionless], range fRatioMin~fRatioMax
    fRatioMin       : REAL := 0.01;           // 比率下限 [无量纲]，必须 > 0 / ratio lower bound [dimensionless], must be > 0
    fRatioMax       : REAL := 10.0;           // 比率上限 [无量纲]，必须 > fRatioMin / ratio upper bound [dimensionless], must be > fRatioMin
    fBias           : REAL := 0.0;            // 偏置量 [m3/h]，范围 -1.0E4~1.0E4 / bias [m3/h], range -1.0E4~1.0E4
    fMasterLowLimit : REAL := 1.0;            // 主动流量低限 [m3/h]，范围 0.0~1.0E6 / master flow low limit [m3/h], range 0.0~1.0E6
    fMasterLowSp    : REAL := 0.0;            // 低限以下的安全给定 [m3/h]，范围 fOutMin~fOutMax / safe setpoint below the low limit [m3/h], range fOutMin~fOutMax
    fOutMin         : REAL := 0.0;            // 输出下限 [m3/h] / output lower bound [m3/h]
    fOutMax         : REAL := 100.0;          // 输出上限 [m3/h]，必须 > fOutMin / output upper bound [m3/h], must be > fOutMin
    fRateMax        : REAL := 50.0;           // 输出最大变化率 [m3/h/s]，范围 0.001~1.0E6 / maximum output rate [m3/h/s], range 0.001~1.0E6
    tSampleTime     : TIME := T#100MS;        // 采样周期 [ms]，范围 1~10000 / sample time [ms], range 1~10000
END_VAR
VAR_OUTPUT
    fSlaveSp        : REAL;                   // 从动侧给定 [m3/h] / slave setpoint [m3/h]
    bMasterLow      : BOOL;                   // 主动流量低于低限，给定已切安全值 / master flow below the low limit, setpoint switched
    bRatioClamped   : BOOL;                   // 比率被限幅 / ratio clamped
    bOutClamped     : BOOL;                   // 输出被上下限或斜率限制 / output limited by the bounds or the ramp
    fEffectiveRatio : REAL;                   // 实际生效比率（含限幅）[无量纲] / effective ratio including the clamp [dimensionless]
    eErr            : UDINT;                  // 错误码，0=正常 / error id, 0=ok
    bError          : BOOL;                   // 故障标志，eErr 为故障级时 TRUE / error flag, TRUE on fault-level eErr
    bValid          : BOOL;                   // 给定是否可用 / setpoint valid flag
END_VAR
VAR
    eState          : E_DL_RatioState := eIdle; // 状态机当前态 / current state machine state
    fbTrigReset     : R_TRIG;                 // 复位上升沿实例，本体首部无条件刷新 / reset edge instance, refreshed unconditionally
    fLastSp         : REAL;                   // 上一拍给定（斜率限制基准）[m3/h] / previous setpoint used by the ramp [m3/h]
    fStep           : REAL;                   // 本拍允许的最大变化量 [m3/h] / maximum allowed change in this cycle [m3/h]
    fDtSec          : REAL;                   // 采样周期换算的秒数 [s] / sample time converted to seconds [s]
    fRatioEff       : REAL;                   // 限幅后的生效比率 [无量纲] / effective ratio after clamping [dimensionless]
    fTarget         : REAL;                   // 钳位与限速率前的目标给定 [m3/h] / target setpoint before clamping and ramping [m3/h]
    bNonFin         : BOOL;                   // 输入非有限判定标志 / non-finite input flag
    nDtMs           : DINT;                   // 采样周期毫秒整数 [ms] / sample time in integer milliseconds [ms]
END_VAR
VAR CONSTANT
    DL_RTO_RATIO_EPS : REAL := 1.0E-6;        // 比率判零容差 [无量纲] / ratio zero tolerance [dimensionless]
    DL_RTO_RATE_MIN  : REAL := 0.001;         // 变化率下限 [m3/h/s] / rate lower bound [m3/h/s]
    DL_RTO_RATE_MAX  : REAL := 1.0E6;         // 变化率上限 [m3/h/s] / rate upper bound [m3/h/s]
    DL_RTO_DT_MAX    : TIME := T#10S;         // 采样周期上限 [ms] / sample time upper bound [ms]
    DL_RTO_DT_MIN    : TIME := T#1MS;         // 采样周期下限 [ms] / sample time lower bound [ms]
    DL_FLOAT_EPS     : REAL := 1.0E-6;        // 浮点判等容差 [无量纲] / float equality tolerance [dimensionless]
    DL_RTO_MS_PER_S  : REAL := 1000.0;        // 毫秒到秒的换算因子 [ms/s] / milliseconds per second [ms/s]
    DL_RTO_INF_GUARD : REAL := 1.0E38;        // 非有限幅值判定阈值 [无量纲] / non-finite magnitude guard [dimensionless]
    DL_RTO_ZERO      : REAL := 0.0;           // 零值常量，避免裸字面量 [无量纲] / zero constant, avoids a bare literal [dimensionless]
END_VAR

// 段 1｜边沿实例无条件周期刷新（红线：严禁放入条件分支）/ segment 1, unconditional edge refresh
fbTrigReset(CLK := bReset);

// 段 2｜输出与错误状态预置（fSlaveSp 不预置，故障时须保持末次有效值）/ segment 2, preset outputs except the held setpoint
eErr := 0;                                    // 预置无错误 / preset no error
bError := FALSE;                              // 预置无故障 / preset no fault
bValid := FALSE;                              // 预置不可用 / preset invalid
bMasterLow := FALSE;                          // 预置非低限态 / preset not in the master-low state
bRatioClamped := FALSE;                       // 预置比率未限幅 / preset ratio not clamped
bOutClamped := FALSE;                         // 预置输出未限幅 / preset output not clamped

// 段 3｜输入非有限闸：给定保持末次有效（切 0 会直接停料）/ segment 3, non-finite gate
bNonFin := (fMasterFlow <> fMasterFlow) OR (fMasterFlow > DL_RTO_INF_GUARD) OR (fMasterFlow < -DL_RTO_INF_GUARD)
        OR (fRatio <> fRatio) OR (fBias <> fBias)
        OR (fRatioMin <> fRatioMin) OR (fRatioMax <> fRatioMax)
        OR (fOutMin <> fOutMin) OR (fOutMax <> fOutMax)
        OR (fMasterLowLimit <> fMasterLowLimit) OR (fMasterLowSp <> fMasterLowSp); // 非有限判定 / non-finite detection
IF bNonFin THEN
    eErr := 16#0002_2810;                     // 输入非有限故障码 / non-finite input fault id
    bError := TRUE;                           // 置故障标志 / raise the error flag
    eState := eFault;         // 落故障态 / enter the fault state
    fSlaveSp := fLastSp;                      // 给定保持末次有效值 / hold the last valid setpoint
    RETURN;                                   // 故障级提前返回 / early return on fault
END_IF

// 段 4｜限值区间自洽闸（区间不存在即故障，比参数越界更危险）/ segment 4, interval consistency gate
IF (fRatioMin <= DL_RTO_RATIO_EPS) OR (fRatioMax <= fRatioMin) THEN
    eErr := 16#0002_2811;                     // 比率域自相矛盾故障码 / ratio domain contradiction fault id
    bError := TRUE;                           // 置故障标志 / raise the error flag
    eState := eFault;         // 落故障态 / enter the fault state
    fSlaveSp := fLastSp;                      // 保持末值 / hold the last value
    RETURN;                                   // 故障级提前返回 / early return on fault
END_IF
IF fOutMax <= fOutMin THEN
    eErr := 16#0002_2811;                     // 输出域自相矛盾，同一语义复用同一故障码 / output domain contradiction, same fault id
    bError := TRUE;                           // 置故障标志 / raise the error flag
    eState := eFault;         // 落故障态 / enter the fault state
    fSlaveSp := fLastSp;                      // 保持末值 / hold the last value
    RETURN;                                   // 故障级提前返回 / early return on fault
END_IF

// 段 5｜斜率与采样参数闸（参数非法则斜率律不可信）/ segment 5, rate and sample gate
IF (fRateMax < DL_RTO_RATE_MIN) OR (fRateMax > DL_RTO_RATE_MAX)
   OR (tSampleTime < DL_RTO_DT_MIN) OR (tSampleTime > DL_RTO_DT_MAX) THEN
    eErr := 16#0002_2810;                     // 斜率或采样参数非法故障码 / rate or sample parameter fault id
    bError := TRUE;                           // 置故障标志 / raise the error flag
    eState := eFault;         // 落故障态 / enter the fault state
    fSlaveSp := fLastSp;                      // 给定保持末次有效值 / hold the last valid setpoint
    RETURN;                                   // 故障级提前返回 / early return on fault
END_IF

// 段 6｜斜率步长（首拍 fLastSp 未建立时 fStep = 0，绝不用 0 除）/ segment 6, ramp step
nDtMs := TIME_TO_DINT(tSampleTime);           // 采样周期显式取整数毫秒 / take the sample time in integer milliseconds
fDtSec := DINT_TO_REAL(nDtMs) / DL_RTO_MS_PER_S; // 换算为秒，除子为常量非零 [s] / convert to seconds, the divisor is a nonzero constant [s]
IF fDtSec <= DL_RTO_ZERO THEN
    fStep := DL_RTO_ZERO;                     // 首拍或非法周期：不突变 / first scan or illegal period, no step at all
ELSE
    fStep := fRateMax * fDtSec;               // 本拍允许的最大变化量 [m3/h] / maximum allowed change in this cycle [m3/h]
END_IF

// 段 7｜复位沿清限幅锁存与斜率状态（不改变状态机态）/ segment 7, reset edge clears the latches
IF fbTrigReset.Q THEN
    fLastSp := MIN(MAX(fLastSp, fOutMin), fOutMax); // 复位把基准拉回合法域 / pull the ramp reference back into the legal domain
    bRatioClamped := FALSE;                   // 清比率限幅锁存 / clear the ratio clamp latch
    bOutClamped := FALSE;                     // 清输出限幅锁存 / clear the output clamp latch
END_IF

// 段 8｜失能无条件回 eIdle / segment 8, disabled forces eIdle
IF NOT bEnable THEN
    eState := eIdle;          // 失能回空闲态 / return to idle when disabled
END_IF

// 段 9｜比率限幅（越窗是待调整，只置信息码）/ segment 9, ratio clamp
fRatioEff := fRatio;                          // 取入参副本 / copy the input
IF fRatioEff > fRatioMax THEN
    fRatioEff := fRatioMax;                   // 越上限钳位 / clamp at the upper bound
    bRatioClamped := TRUE;                    // 标记比率限幅 / flag the ratio clamp
    eErr := 16#0002_2801;                     // 信息级：比率被限幅 / info level, the ratio was clamped
ELSIF fRatioEff < fRatioMin THEN
    fRatioEff := fRatioMin;                   // 越下限钳位 / clamp at the lower bound
    bRatioClamped := TRUE;                    // 标记比率限幅 / flag the ratio clamp
    eErr := 16#0002_2801;                     // 同一业务语义复用同一信息码 / the same semantics reuses the same info id
END_IF
fEffectiveRatio := fRatioEff;                 // 发布生效比率 / publish the effective ratio

// 段 10｜状态机（含 ELSE 兜底）/ segment 10, state machine with ELSE fallback
CASE eState OF
    eIdle:
        fSlaveSp := fOutMin;                  // 空闲态输出限幅下限，不按比例算 / idle outputs the lower bound, no ratio computation
        fLastSp := fOutMin;                   // 斜率基准同步，避免使能首拍跳变 / sync the ramp reference to avoid a jump on enable
        IF bEnable THEN
            eState := eRunning; // 使能即进入运行态 / enabling enters the running state
        END_IF

    eRunning:
        IF fMasterFlow < fMasterLowLimit THEN
            fTarget := fMasterLowSp;          // 低限以下切安全给定，不按比例算 / below the low limit switch to the safe setpoint
            bMasterLow := TRUE;               // 发布低限标志 / publish the master-low flag
            eErr := 16#0002_2801;             // 信息级：主动流量低于低限已切安全给定 / info level, the safe setpoint was applied
            eState := eMasterLow; // 迁移到低限态 / move to the master-low state
        ELSE
            fTarget := fMasterFlow * fRatioEff + fBias; // 比值律：从动给定 = 主动 × 比率 + 偏置 / ratio law
        END_IF

    eMasterLow:
        fTarget := fMasterLowSp;              // 低限态保持安全给定 / hold the safe setpoint in the master-low state
        bMasterLow := TRUE;                   // 持续发布低限标志 / keep publishing the master-low flag
        IF fMasterFlow >= fMasterLowLimit THEN
            eState := eRunning; // 主动流量恢复即回运行态 / return to running once the master recovers
        END_IF

    eFault:
        fTarget := fLastSp;                   // 故障态目标即末次值，不再跟踪 / the fault state targets the last value, no tracking
        bValid := FALSE;                      // 故障态给定不可用 / the setpoint is not usable in the fault state

ELSE
    eErr := 16#0002_2812;                     // 故障级：非法状态兜底 / fault level, illegal state fallback
    bError := TRUE;                           // 置故障标志 / raise the error flag
    eState := eIdle;          // 回空闲态 / fall back to idle
    fTarget := fLastSp;                       // 保持末值，不产生跳变 / hold the last value, no jump
END_CASE

// 段 11｜输出双侧钳位（只做单侧是常见缺陷）/ segment 11, two-sided output clamp
IF fTarget > fOutMax THEN
    fTarget := fOutMax;                       // 上限钳位 / clamp at the upper bound
    bOutClamped := TRUE;                      // 标记输出限幅 / flag the output clamp
ELSIF fTarget < fOutMin THEN
    fTarget := fOutMin;                       // 下限钳位 / clamp at the lower bound
    bOutClamped := TRUE;                      // 标记输出限幅 / flag the output clamp
END_IF

// 段 12｜斜率限制（每拍最多变化 fStep）/ segment 12, ramp limiting
IF fStep > DL_RTO_ZERO THEN
    IF fTarget > (fLastSp + fStep) THEN
        fTarget := fLastSp + fStep;           // 正向每拍限幅 / limit the positive step per cycle
        bOutClamped := TRUE;                  // 标记斜率限制 / flag the ramp limit
    ELSIF fTarget < (fLastSp - fStep) THEN
        fTarget := fLastSp - fStep;           // 负向每拍限幅 / limit the negative step per cycle
        bOutClamped := TRUE;                  // 标记斜率限制 / flag the ramp limit
    END_IF
END_IF

// 段 13｜发布给定与状态（无故障时给定可用）/ segment 13, publish the setpoint and the status
fSlaveSp := fTarget;                          // 输出本拍给定 [m3/h] / publish this cycle setpoint [m3/h]
fLastSp := fTarget;                           // 记录为下一拍斜率基准 / remember it as the next ramp reference
IF NOT bError THEN
    bValid := TRUE;                           // 无故障则给定可用 / usable when no fault is present
END_IF
END_FUNCTION_BLOCK

(* ---- FB_DL_RatioStationCalc.st ---- *)
(*
  FB_DL_RatioStationCalc  —  比值站：随动设定 = K×主流量 + 偏置 / Ratio station: K times master flow plus offset
  分类 Category : DL_Algo
  版本 Version  : 1.0.0
  来源 Source   : t2-2-lbp — 比值控制族零检索深化
  溯源 Origin   : clean-room 实现，未复制任何源码行
  功能 Function : 1) 双模式：eRatio（随动 fSetpoint := K×fMaster + fOffset）/
                  eFixed（fSetpoint := fFixedSet）；eMode 落枚举域外 → CASE ELSE → 03AA；
                  2) 主流量非有限（NaN 自反判 / Inf 差值自减判）→ bMasterOk FALSE，
                  强制切固定模式并置信息级 048F；恢复有限自动回比值模式；
                  3) K 组态域钳位 [0.0, 100.0]，钳位发生置信息级 0490；
                  4) 模式变更沿 bModeChg 单拍脉冲（当拍量比较，禁锁存量自指）。
  边界 Boundary : ① 组态闸：fK / fOffset / fFixedSet 非有限 → 03A9 锁存；
                  ② 模式切换 bModeChg 为单拍脉冲：内部 _b* 置位 → 统一出口映射（禁同拍抹除）；
                  ③ 钳位域常量固定，域内无除法，无除零路径；
                  ④ 无 GVL 依赖：纯引脚输入输出，无外部变量引用，无物理 IO 地址。
  依赖 Depends  : 仅 Standard.library（ABS / REAL 算术）
  码表 Error codes（Algo 段 0002，窗口 03A9~03AA / 048F~0490）:
    16#0002_03A9 故障级：组态非有限（fK/fOffset/fFixedSet 任一非有限），锁存至 bReset
    16#0002_03AA 故障级：模式落 CASE ELSE 兜底（非法 eMode），锁存至 bReset
    16#0002_048F 信息级：主流量无效，强制固定模式（恢复有限自动回比值）
    16#0002_0490 信息级：K 已钳位至组态域 [0, 100]
  修订历史 Revision :
    2026-11-19  v1.0.0  R41 首版（批次 3 · 序号 4）
*)

TYPE E_DL_RatioMode :
(
    eRatio := 0,   // 比值模式：随动设定 / Ratio mode, slave setpoint
    eFixed := 10   // 固定模式：固定设定 / Fixed mode, constant setpoint
);
END_TYPE

FUNCTION_BLOCK FB_DL_RatioStationCalc
VAR_INPUT
    fMaster      : REAL := 0.0;       // 主流量 [EU] / Master flow
    fK           : REAL := 1.0;       // 比值系数 [无量纲]，域 [0, 100] 钳位生效 / Ratio factor
    fOffset      : REAL := 0.0;       // 偏置 [EU] / Offset
    fFixedSet    : REAL := 0.0;       // 固定模式设定值 [EU] / Fixed-mode setpoint
    eMode        : E_DL_RatioMode := E_DL_RatioMode.eRatio;  // 模式选择 / Mode select
    bEnable      : BOOL := FALSE;     // 投运使能 [-] / Enable
    bReset       : BOOL := FALSE;     // 复位，上升沿清故障锁存 / Reset edge clears fault latch
END_VAR
VAR_OUTPUT
    fSetpoint    : REAL;              // 随动/固定设定值出口 [EU] / Setpoint outlet
    bMasterOk    : BOOL;              // 主流量有效标志 [-] / Master validity flag
    bModeChg     : BOOL;              // 模式变更单拍脉冲 [-] / Mode change one-shot pulse
    bValid       : BOOL;              // 输出有效标志 / Output valid flag
    bError       : BOOL;              // 故障锁存标志 / Fault latch flag
    nErrId       : UDINT;             // 事件码，0 = 无事件 / Event code
END_VAR
VAR
    rtReset      : R_TRIG;            // 复位沿实例，无条件刷新 / Reset edge instance
    _fKEff       : REAL;              // 钳位后生效比值系数 / Effective clamped factor
    _bMasterFin  : BOOL;              // 主流量有限当拍量 [-] / Master finite current-scan flag
    _eModePrev   : E_DL_RatioMode := E_DL_RatioMode.eRatio;  // 上拍模式快照（变更沿判据）/ Previous mode
    _bModeChgInt : BOOL;              // 模式变更内部脉冲（两段式出口）/ Internal mode-change pulse
    _bFault      : BOOL;              // 故障锁存位（锁存量）/ Latched fault bit
    _uFault      : UDINT;             // 故障码锁存（锁存量）/ Latched fault code
    _uInfo       : UDINT;             // 信息码，每拍重算 / Transient info code
END_VAR
VAR CONSTANT
    DL_RSC_K_MIN : REAL := 0.0;      // 比值系数下限 [无量纲] / Factor lower bound
    DL_RSC_K_MAX : REAL := 100.0;    // 比值系数上限 [无量纲] / Factor upper bound
END_VAR

(* —— 段 0：沿实例无条件周期刷新（禁置于 IF/CASE 内） —— *)
rtReset(CLK := bReset);             // 复位沿（每拍必调）

(* —— 段 1：单拍量预清零（锁存量 _bFault/_uFault 不入清单；脉冲两段式出口） —— *)
_uInfo := 16#0000_0000;             // 信息码每拍重算
bModeChg := FALSE;                  // 模式变更脉冲缺省 FALSE
bValid := FALSE;                    // 有效出口缺省 FALSE
nErrId := 16#0000_0000;             // 事件码缺省无事件
_bModeChgInt := FALSE;              // 内部脉冲清零
fSetpoint := 0.0;                   // 设定值缺省 0

(* —— 段 2：复位沿 + 组态域闸（当拍量判据） —— *)
IF rtReset.Q THEN                   // rtReset.Q = 当拍量
    _bFault := FALSE;               // 清故障锁存位
    _uFault := 16#0000_0000;        // 清故障锁存码
END_IF
IF (fK <> fK) OR (fOffset <> fOffset) OR (fFixedSet <> fFixedSet)
   OR ((fK - fK) <> (fK - fK)) OR ((fOffset - fOffset) <> (fOffset - fOffset))
   OR ((fFixedSet - fFixedSet) <> (fFixedSet - fFixedSet)) THEN
    _uFault := 16#0002_03A9;        // 故障级：组态非有限
    _bFault := TRUE;
END_IF

(* —— 段 3：K 钳位与主流量有效性（当拍量判据） —— *)
_fKEff := fK;                       // 生效系数初值
IF _fKEff < DL_RSC_K_MIN THEN
    _fKEff := DL_RSC_K_MIN;         // 下界钳位
    _uInfo := 16#0002_0490;         // 信息级：K 已钳位
ELSIF _fKEff > DL_RSC_K_MAX THEN
    _fKEff := DL_RSC_K_MAX;         // 上界钳位
    _uInfo := 16#0002_0490;         // 信息级：K 已钳位
END_IF
_bMasterFin := (fMaster = fMaster) AND ((fMaster - fMaster) = (fMaster - fMaster));
                                    // 主流量有限判定：NaN 自反取反 AND Inf 差值自减取反
bMasterOk := _bMasterFin;           // 有效性出口镜像

(* —— 段 4：模式变更沿（当拍量比较，禁锁存量自指） —— *)
IF eMode <> _eModePrev THEN
    _bModeChgInt := TRUE;           // 内部脉冲置位（出口段统一映射）
END_IF
_eModePrev := eMode;                // 模式快照推进（段末统一写口径前移）

(* —— 段 5：设定值仲裁（CASE 全覆盖 + ELSE 兜底） —— *)
CASE eMode OF

E_DL_RatioMode.eRatio:
    IF _bMasterFin THEN
        fSetpoint := fMaster * _fKEff + fOffset;    // 比值随动设定
    ELSE
        fSetpoint := fFixedSet;     // 主流量无效：退固定模式
        _uInfo := 16#0002_048F;     // 信息级：无效退固定
    END_IF

E_DL_RatioMode.eFixed:
    fSetpoint := fFixedSet;         // 固定设定直通

ELSE
    _uFault := 16#0002_03AA;        // 故障级：非法模式兜底
    _bFault := TRUE;
    fSetpoint := 0.0;               // 安全侧归零

END_CASE

(* —— 段 6：出口单点映射（脉冲两段式：内部 _b* → 统一出口；锁存码回放） —— *)
IF _bModeChgInt THEN
    bModeChg := TRUE;               // 模式变更脉冲单拍出口
END_IF
bValid := (NOT _bFault) AND bEnable;    // 有效出口
IF _bFault THEN
    nErrId := _uFault;              // 故障锁存码回放
    bValid := FALSE;                // 故障期强制 FALSE（安全侧）
ELSE
    nErrId := _uInfo;               // 信息码
END_IF
bError := _bFault;                  // 故障标志与锁存位同源

END_FUNCTION_BLOCK

(* ---- FB_DL_RelayAutoTune.st ---- *)
(*
  组件名 Component   : FB_DL_RelayAutoTune
  子库 Sublibrary    : DL_Algo
  版本 Version       : 1.0.0
  兼容性 Platform    : CODESYS 3.5 / TwinCAT 3 / 汇川 InoProShop / Machine Expert（仅 Standard.library）
  功能 Function      : 继电器反馈法 PID 自整定（只出参数、不闭环）：
                       1) 继电器试验：被控量低于（设定值-迟滞）输出继电器上限，高于
                       （设定值+迟滞）输出继电器下限，形成极限环；
                       2) 极限环测量：继电器同向切换沿间隔 = 振荡周期 Tu，切换沿间
                       被控量峰谷差 / 2 = 振荡幅值 a；
                       3) 临界增益 Ku = 4d / (π·a)（幅值近零前置拦截，不进入除法）；
                       4) Ziegler-Nichols 公开判据初值：Kp = 0.6Ku，Ti = 0.5Tu，Td = 0.125Tu；
                       5) 连续 3 个完整振荡周期取均值后才出参数，试验无切换超时即判故障。
  边界 Boundary      : ① 本件只出初值参数，不接管回路闭环（上层自选时机装载）；
                       ② 振幅近零（a < 容差）→ 故障锁存：被控量不振荡，Ku 无意义；
                       ③ 幅值测量在切换沿间闭环刷新，峰谷快照在切换沿复归；
                       ④ 试验超时计时以切换沿重启（bGuardHold 单拍驻留，见段 0 注释）；
                       ⑤ 故障锁存解除唯一路径 = bReset 上升沿（输入引脚，恒可达）；
                       ⑥ 无全局变量引用、无外部变量声明、无物理地址寻址。
  依赖 Depends       : Standard.library（R_TRIG / TON）
  溯源 Origin        : 道莅自研 clean-room（参考 t2-5-modpid 参数域与公开 Ziegler-Nichols
                       判据文献语义，零代码行复制）
  码位 Code          : 16#02_3_8D
  码表 Error codes（Algo 格 02_3_8D，单轨：故障 0x038D / 信息 0x028D）:
    16#0002_038D 故障级：试验非法（无切换超时 / 振幅近零 / 组态非法 / 输入非有限），
                 锁存至 bReset 上升沿
    16#0002_028D 信息级：整定完成沿（参数写定拍，锁存至 bReset）
  修订历史 Revision  :
    2026-11-19  v1.0.0  R44 首版（批次 1 · 序号 3）
*)

TYPE E_DL_RatState :
(
    eIdle  := 0,    // 空闲：等启动沿 / Idle, waiting start edge
    eTune  := 10,   // 试验：继电器极限环运行中 / Tuning, relay limit cycle running
    eDone  := 20,   // 完成：参数驻留待装载 / Done, parameters held
    eFault := 90    // 故障：试验非法锁存 / Fault, latched
);
END_TYPE

FUNCTION_BLOCK FB_DL_RelayAutoTune
VAR_INPUT
    bStartCmd  : BOOL;                     // 启动沿（试验以上升沿承载）[-] / Start command edge
    bReset     : BOOL;                     // 上升沿清故障与完成结果 [-] / Reset edge
    fPv        : REAL;                     // 被控量 [工程单位] / Process variable
    fBiasPv    : REAL;                     // 继电器中心（目标值）[工程单位] / Relay bias point
    fHysteresis: REAL := 1.0;              // 继电器迟滞半宽 [工程单位] / Relay hysteresis half band
    fRelayHi   : REAL := 100.0;            // 继电器上限输出 [%] / Relay high output
    fRelayLo   : REAL := 0.0;              // 继电器下限输出 [%] / Relay low output
    fRelayAmp  : REAL := 5.0;              // 继电器幅值 d = (上限-下限)/2 [%] / Relay amplitude d
    tGuardTo   : TIME := T#120S;           // 无切换超时 [毫秒]，以切换沿重启 / No-switch timeout
    tCycle     : TIME := T#10MS;           // 扫描周期 [毫秒] / Scan cycle time
END_VAR
VAR_OUTPUT
    fRelayOut  : REAL;                     // 试验期继电器输出 [%]，空闲相 0 / Relay output during test
    bTuning    : BOOL;                     // 试验进行中标志 [-] / Tuning active flag
    bDone      : BOOL;                     // 整定完成锁存标志 [-] / Tune done latch
    fKpInit    : REAL;                     // Z-N 初值比例增益 [无量纲] / ZN initial Kp
    fTiInit    : REAL;                     // Z-N 初值积分时间 [秒] / ZN initial Ti
    fTdInit    : REAL;                     // Z-N 初值微分时间 [秒] / ZN initial Td
    fTuMeas    : REAL;                     // 实测振荡周期 [秒] / Measured ultimate period
    fKuMeas    : REAL;                     // 实测临界增益 [无量纲] / Measured ultimate gain
    eState     : E_DL_RatState;            // 状态出口，段尾单点映射 / State outlet
    bError     : BOOL;                     // 故障锁存标志 [-] / Fault latch flag
    uErrId     : UDINT;                    // 事件码，0 = 无事件 / Event code
END_VAR
VAR
    rtStart    : R_TRIG;                   // 启动沿实例，段 0 无条件刷新 / Start edge
    rtReset    : R_TRIG;                   // 复位沿实例，段 0 无条件刷新 / Reset edge
    rtRelayHi  : R_TRIG;                   // 继电器上沿实例，段 0 无条件刷新 / Relay rising edge
    rtRelayLo  : R_TRIG;                   // 继电器下沿实例，段 0 无条件刷新 / Relay falling edge
    tonGuardTo : TON;                      // 无切换超时（专用超时件（R228A 合法豁免命名）） / No-switch timeout
    _eState    : E_DL_RatState := E_DL_RatState.eIdle;   // 内部相位（CASE 唯一写入目标） / Internal phase
    _bRelHi    : BOOL;                     // 继电器上电平（迟滞内部态）[-] / Relay high level state
    _fPk       : REAL;                     // 本周期峰快照 [工程单位] / Peak snapshot
    _fVl       : REAL;                     // 本周期谷快照 [工程单位] / Valley snapshot
    _fAmpSum   : REAL;                     // 幅值累加 [工程单位] / Amplitude accumulator
    _fTuSum    : REAL;                     // 周期累加 [秒] / Period accumulator
    _fTuCur    : REAL;                     // 本周期秒计 [秒] / Current period seconds
    _nCyc      : DINT;                     // 切换沿计数 [个] / Switch edge count
    _fAmpAvg   : REAL;                     // 幅值均值 [工程单位] / Amplitude average
    _bGuardHold: BOOL;                     // 超时重启驻留（切换沿置位，下拍段 1 清除）[-] / Guard restart hold
    _bFault    : BOOL;                     // 故障锁存位（锁存量） / Latched fault bit
    _uFault    : UDINT;                    // 故障码锁存（锁存量） / Latched fault code
    _bCfgBad   : BOOL;                     // 组态非法当拍量 [-] / Config illegal flag
    _fCyS      : REAL;                     // 扫描周期秒值 [秒] / Cycle seconds
END_VAR
VAR CONSTANT
    DL_CYC_REQ  : INT   := 3;              // 取均值所需完整周期数 [个] / Cycles to average
    DL_EDGES_REQ: DINT  := 6;              // 完整周期对应切换沿数 = 2 × 周期数 [个] / Required edges
    DL_ZN_KP    : REAL  := 0.6;            // Z-N 比例判据系数 [无量纲] / ZN Kp coefficient
    DL_ZN_TI    : REAL  := 0.5;            // Z-N 积分判据系数 [无量纲] / ZN Ti coefficient
    DL_ZN_TD    : REAL  := 0.125;          // Z-N 微分判据系数 [无量纲] / ZN Td coefficient
    DL_PI       : REAL  := 3.14159265;     // 圆周率 [无量纲] / Pi constant
    DL_AMP_MIN  : REAL  := 1.0E-6;         // 幅值近零判据 [工程单位] / Amplitude near-zero threshold
    DL_AMP_FACT : REAL  := 4.0;            // Ku = 4d/(π·a) 分子系数 [无量纲] / Ku numerator factor
    DL_HALF     : REAL  := 0.5;            // 峰谷差折半系数 [无量纲] / Half factor
    DL_KU_MIN   : REAL  := 1.0E-6;         // 临界增益下限护栏 [无量纲] / Ku floor
    DL_ABS_MAX  : REAL  := 1.0E30;         // 有限值判定上界 [工程单位] / Finite bound
    DL_ZERO     : REAL  := 0.0;            // 零常量 [工程单位] / Zero constant
    DL_TWO      : REAL  := 2.0;            // 二常量 [无量纲] / Two constant
    DL_MS_PER_S : REAL  := 1000.0;         // 毫秒 → 秒换算系数 [毫秒/秒] / Milliseconds per second
END_VAR

(* —— 段 0｜沿与定时器每拍无条件刷新（禁置于 IF/CASE 内；bGuardHold 切换沿置位、
        下拍段 1 清除，tonGuardTo 以此实现逐切换沿重启，IN 两拍一断合法复位） —— *)
rtStart  (CLK := bStartCmd);
rtReset  (CLK := bReset);
rtRelayHi(CLK := _bRelHi);
rtRelayLo(CLK := NOT _bRelHi);
tonGuardTo(IN := (_eState = E_DL_RatState.eTune) AND (NOT _bGuardHold), PT := tGuardTo);

(* —— 段 1｜瞬时量预清零（锁存量 _bFault/_uFault/bDone/_bRelHi 不入清单） —— *)
_bGuardHold := FALSE;                    // 超时重启驻留只驻留一拍
_bCfgBad    := FALSE;
uErrId      := 16#0000_0000;
_fCyS       := TIME_TO_REAL(tCycle) / DL_MS_PER_S;

(* —— 段 2｜复位沿：故障、完成结果、测量累计一次性清干净 —— *)
IF rtReset.Q THEN
    _bFault  := FALSE;
    _uFault  := 16#0000_0000;
    bDone    := FALSE;
    _nCyc    := 0;
    _fAmpSum := DL_ZERO;
    _fTuSum  := DL_ZERO;
    _fTuCur  := DL_ZERO;
    IF _eState = E_DL_RatState.eFault THEN
        _eState := E_DL_RatState.eIdle;  // eFault 迁出唯一属主 = rtReset.Q（可达）
    END_IF
END_IF

(* —— 段 3｜组态闸：迟滞/幅值/周期域与非有限值前置拦截 —— *)
IF (fHysteresis <= DL_ZERO) OR (fRelayAmp <= DL_ZERO) OR (tGuardTo = T#0S) OR (tCycle = T#0S)
   OR (fPv <> fPv) OR (fBiasPv <> fBiasPv) OR (fHysteresis > DL_ABS_MAX) THEN
    _bCfgBad := TRUE;
END_IF

(* —— 段 4｜主状态机：四态全覆盖 + ELSE 兜底 —— *)
CASE _eState OF

E_DL_RatState.eIdle:
    fRelayOut := DL_ZERO;                // 空闲继电器输出回零（安全侧）
    IF _bFault THEN
        bError := TRUE;                  // 故障锁存回放（R189）
    END_IF
    IF rtStart.Q AND (NOT _bFault) AND (NOT _bCfgBad) THEN
        _bRelHi  := FALSE;               // 继电器从下限起振
        _fPk     := fPv;                 // 峰谷快照初始化
        _fVl     := fPv;
        _fTuCur  := DL_ZERO;
        _nCyc    := 0;
        _fAmpSum := DL_ZERO;
        _fTuSum  := DL_ZERO;
        bDone    := FALSE;
        _eState  := E_DL_RatState.eTune;
    ELSIF rtStart.Q AND (_bCfgBad OR _bFault) THEN
        _bFault := TRUE;                 // 带病启动拒绝
        _uFault := 16#0002_038D;
        bError  := TRUE;
        _eState := E_DL_RatState.eFault;
    END_IF

E_DL_RatState.eTune:
    bTuning := TRUE;
    (* 继电器迟滞逻辑：低于中心-迟滞输出上限，高于中心+迟滞输出下限 *)
    IF (NOT _bRelHi) AND (fPv < fBiasPv - fHysteresis) THEN
        _bRelHi := TRUE;
    ELSIF _bRelHi AND (fPv > fBiasPv + fHysteresis) THEN
        _bRelHi := FALSE;
    END_IF
    IF _bRelHi THEN
        fRelayOut := fRelayHi;
    ELSE
        fRelayOut := fRelayLo;
    END_IF

    (* 峰谷跟踪与周期秒计 *)
    IF fPv > _fPk THEN
        _fPk := fPv;
    END_IF
    IF fPv < _fVl THEN
        _fVl := fPv;
    END_IF
    _fTuCur := _fTuCur + _fCyS;

    IF rtRelayHi.Q OR rtRelayLo.Q THEN
        (* 切换沿：相邻沿间隔 × 2 = 一个完整振荡周期，幅值按沿取样 *)
        _fTuSum := _fTuSum + _fTuCur * DL_TWO;
        _fAmpSum := _fAmpSum + (_fPk - _fVl) * DL_HALF;
        _fTuCur  := DL_ZERO;
        _fPk     := fPv;                 // 峰谷快照按沿复归
        _fVl     := fPv;
        _bGuardHold := TRUE;             // 超时计时重启驻留（下拍断 IN）
        _nCyc := _nCyc + 1;
        IF _nCyc >= DL_EDGES_REQ THEN
            (* 收口：均值 → 临界参数 → Z-N 公开判据初值（除数 = 沿数 > 0 已由闸保证） *)
            _fAmpAvg := _fAmpSum / DINT_TO_REAL(_nCyc);
            IF _fAmpAvg < DL_AMP_MIN THEN
                _bFault := TRUE;         // 振幅近零：Ku 无意义
                _uFault := 16#0002_038D;
                bError  := TRUE;
                _eState := E_DL_RatState.eFault;
            ELSE
                fTuMeas := _fTuSum / DINT_TO_REAL(_nCyc);
                fKuMeas := (DL_AMP_FACT * fRelayAmp) / (DL_PI * _fAmpAvg);
                IF fKuMeas < DL_KU_MIN THEN
                    fKuMeas := DL_KU_MIN;            // 临界增益下限钳位
                END_IF
                fKpInit := DL_ZN_KP * fKuMeas;
                fTiInit := DL_ZN_TI * fTuMeas;
                fTdInit := DL_ZN_TD * fTuMeas;
                uErrId  := 16#0002_028D;     // 信息级：整定完成沿（锁存至复位）
                bDone   := TRUE;
                bTuning := FALSE;
                _eState := E_DL_RatState.eDone;
            END_IF
        END_IF
    END_IF

    IF tonGuardTo.Q THEN
        _bFault := TRUE;                 // 无切换超时：过程不振荡
        _uFault := 16#0002_038D;
        bError  := TRUE;
        bTuning := FALSE;
        fRelayOut := DL_ZERO;            // 安全侧回零
        _eState := E_DL_RatState.eFault;
    END_IF

E_DL_RatState.eDone:
    bTuning := FALSE;
    fRelayOut := DL_ZERO;                // 完成相继电器输出回零
    IF NOT bStartCmd THEN
        _eState := E_DL_RatState.eIdle;  // 启动指令撤销：回空闲（结果锁存保留）
    END_IF

E_DL_RatState.eFault:
    bTuning := FALSE;
    fRelayOut := DL_ZERO;
    bError := TRUE;
    ;                                    // 故障相驻留：只认复位沿（段 2 承载迁出）

ELSE
    _bFault := TRUE;                     // 兜底：非法相位锁存
    _uFault := 16#0002_038D;
    bError  := TRUE;
    _eState := E_DL_RatState.eFault;
END_CASE

(* —— 段 5｜状态出口单点映射 —— *)
eState := _eState;
END_FUNCTION_BLOCK
